(* IEC 61131-3 sources: 2026_Projet_YGO_ExcavatriceDragage/TOOLS/TEST_AUTO_CI/RESULTS/H_TREUILS_BENNE/reports (part 2) *)

(* ---- FB_BucketCloseThreshold_test.st ---- *)
(* =======================================================================
   🧪 FB_BucketCloseThreshold — seuil IHM d'ouverture benne (T262 phase B, C4)
   ───────────────────────────────────────────────────────────────────────
   Périmètre STRICT : le FB de décision en BOÎTE NOIRE. Il dérive du réglage
   IHM `ExtractionStartOpening_Pct` une DISTANCE de fermeture équivalente et
   un signal `Reached`. Il ne lit ni GVL, ni FB_Bucket, ni le cycle : aucun
   consommateur n'est testé ici (PRG_04 / FB_Bucket / FB_CycleSemiAuto
   relèvent de l'essai CODESYS et des gates mécaniques).

   ── Propriété cardinale (AC2 du contrat T262-PHASE-B) ──────────────────
   À ThresholdPct = 0, la branche est INACTIVE PAR CONSTRUCTION : `Reached`
   reste FALSE sur TOUTE la table Delta x géométrie. C'est ce qui rend la
   non-régression du comportement historique indépendante d'un MAX.

   ── Conventions ────────────────────────────────────────────────────────
   1) 1 appel `fb(...)` = 1 scan. Le FB est PUR (aucun état, aucun timer).
   2) ⚠️ Aucune assertion dans une boucle FOR/WHILE : ce build STruCpp
      SUPPRIME silencieusement les ASSERT_* du corps d'une boucle (vérifié
      dans le C++ généré). Tous les balayages sont DÉROULÉS.
   3) Tolérance 1e-6 : REAL en simple précision, littéral ST lu en double.
      Les distances attendues (p x 0,15 m) sont exactes à 1e-6 près.

   ── Géométrie de référence (valeurs persistées GVL_PERSISTENT) ─────────
   OffsetOpenM = 0,0 m · OffsetCloseM = 15,0 m · débattement = 15,0 m
   ⇒ distance équivalente = p % x 15,0 m = p x 0,15 m

   Références : DOC/WFLOW/AUDITS/DESIGN/CHALLENGE_T262_PHASE_B_SEUIL_BENNE_2026-09-21.md
                DOC/WFLOW/CONTRACTS/TASK_CONTRACT_T262_PHASE_B_BUCKET_OPENING_THRESHOLD.yaml
   ======================================================================= *)

SETUP
VAR
    FB : FB_BucketCloseThreshold;
END_VAR
END_SETUP

(* ── Groupe A · Branche INACTIVE à 0 % (AC2, AC4) ─────────────────────── *)

TEST 'TC-T262B-001 seuil 0 % : Reached FAUX sur toute la table Delta x geometrie'
    (* Balayage DEROULE. Geometrie nominale 0,0 / 15,0 m ; qualification pleine. *)
    FB.ThresholdPct := 0;
    FB.OffsetOpenM := 0.0;
    FB.OffsetCloseM := 15.0;
    FB.MeasureValid := TRUE;
    FB.IsIntermediate := TRUE;

    FB.DeltaPosition_M := 0.0;   FB();
    ASSERT_FALSE(FB.Reached, '0 % : benne ouverte (Delta = 0,0) -> Reached FAUX');
    ASSERT_FALSE(FB.Active,  '0 % : branche seuil INACTIVE');

    FB.DeltaPosition_M := 7.5;   FB();
    ASSERT_FALSE(FB.Reached, '0 % : mi-course (Delta = 7,5) -> Reached FAUX');

    FB.DeltaPosition_M := 13.0;  FB();
    ASSERT_FALSE(FB.Reached, '0 % : au seuil de la tolerance historique -> Reached FAUX');

    FB.DeltaPosition_M := 14.0;  FB();
    ASSERT_FALSE(FB.Reached, '0 % : benne fermee (Delta = 14,0) -> Reached FAUX');

    FB.DeltaPosition_M := 15.0;  FB();
    ASSERT_FALSE(FB.Reached, '0 % : sur la reference fermee -> Reached FAUX (0 % n autorise RIEN)');

    FB.DeltaPosition_M := 16.0;  FB();
    ASSERT_FALSE(FB.Reached, '0 % : sur-fermeture -> Reached FAUX');

    (* Geometrie derivee : la branche doit rester inerte quelle que soit la geometrie. *)
    FB.OffsetOpenM := -1.0;
    FB.OffsetCloseM := 20.0;
    FB.DeltaPosition_M := 19.5;  FB();
    ASSERT_FALSE(FB.Reached, '0 % : autre geometrie (debattement 21,0) -> Reached FAUX');
    ASSERT_NEAR(FB.Distance_M, 0.0, 0.000001, '0 % : distance equivalente EXACTEMENT 0,0 m');
END_TEST

TEST 'TC-T262B-002 distance equivalente : 0,15 m par pourcent (geometrie persistee)'
    (* Balayage DEROULE de p = 0 a 20 : la distance est p x 0,15 m. *)
    FB.OffsetOpenM := 0.0;
    FB.OffsetCloseM := 15.0;
    FB.MeasureValid := TRUE;
    FB.IsIntermediate := TRUE;
    FB.DeltaPosition_M := 0.0;

    FB.ThresholdPct := 0;  FB();  ASSERT_NEAR(FB.Distance_M, 0.0,  0.000001, 'p=0  -> 0,00 m');
    FB.ThresholdPct := 1;  FB();  ASSERT_NEAR(FB.Distance_M, 0.15, 0.000001, 'p=1  -> 0,15 m');
    FB.ThresholdPct := 2;  FB();  ASSERT_NEAR(FB.Distance_M, 0.30, 0.000001, 'p=2  -> 0,30 m');
    FB.ThresholdPct := 3;  FB();  ASSERT_NEAR(FB.Distance_M, 0.45, 0.000001, 'p=3  -> 0,45 m');
    FB.ThresholdPct := 4;  FB();  ASSERT_NEAR(FB.Distance_M, 0.60, 0.000001, 'p=4  -> 0,60 m');
    FB.ThresholdPct := 5;  FB();  ASSERT_NEAR(FB.Distance_M, 0.75, 0.000001, 'p=5  -> 0,75 m');
    FB.ThresholdPct := 6;  FB();  ASSERT_NEAR(FB.Distance_M, 0.90, 0.000001, 'p=6  -> 0,90 m');
    FB.ThresholdPct := 7;  FB();  ASSERT_NEAR(FB.Distance_M, 1.05, 0.000001, 'p=7  -> 1,05 m');
    FB.ThresholdPct := 8;  FB();  ASSERT_NEAR(FB.Distance_M, 1.20, 0.000001, 'p=8  -> 1,20 m (= plancher historique)');
    FB.ThresholdPct := 9;  FB();  ASSERT_NEAR(FB.Distance_M, 1.35, 0.000001, 'p=9  -> 1,35 m');
    FB.ThresholdPct := 10; FB();  ASSERT_NEAR(FB.Distance_M, 1.50, 0.000001, 'p=10 -> 1,50 m');
    FB.ThresholdPct := 13; FB();  ASSERT_NEAR(FB.Distance_M, 1.95, 0.000001, 'p=13 -> 1,95 m');
    FB.ThresholdPct := 14; FB();  ASSERT_NEAR(FB.Distance_M, 2.10, 0.000001, 'p=14 -> 2,10 m (au-dela de la tolerance 2,0)');
    FB.ThresholdPct := 19; FB();  ASSERT_NEAR(FB.Distance_M, 2.85, 0.000001, 'p=19 -> 2,85 m');
    FB.ThresholdPct := 20; FB();  ASSERT_NEAR(FB.Distance_M, 3.00, 0.000001, 'p=20 -> 3,00 m (borne haute)');
END_TEST

(* ── Groupe B · Saturation de la borne 0..20 (AC1) ────────────────────── *)

TEST 'TC-T262B-003 borne basse : seuil negatif ramene a 0 (branche INACTIVE)'
    FB.ThresholdPct := -1;
    FB.OffsetOpenM := 0.0;
    FB.OffsetCloseM := 15.0;
    FB.MeasureValid := TRUE;
    FB.IsIntermediate := TRUE;
    FB.DeltaPosition_M := 14.9;
    FB();
    ASSERT_FALSE(FB.Active, 'Seuil -1 % : branche INACTIVE');
    ASSERT_FALSE(FB.Reached, 'Seuil -1 % : Reached FAUX (aucune autorisation sur saisie hors plage)');
    ASSERT_NEAR(FB.Distance_M, 0.0, 0.000001, 'Seuil -1 % : distance ramenee a 0,0 m');
END_TEST

TEST 'TC-T262B-004 borne haute : seuil 21 ramene a 20 (jamais au-dela)'
    FB.ThresholdPct := 21;
    FB.OffsetOpenM := 0.0;
    FB.OffsetCloseM := 15.0;
    FB.MeasureValid := TRUE;
    FB.IsIntermediate := TRUE;
    FB.DeltaPosition_M := 11.5;   (* ouverture 23,3 % : hors de la plage autorisee *)
    FB();
    ASSERT_NEAR(FB.Distance_M, 3.00, 0.000001, 'Seuil 21 % : distance CLAMPEE a 3,00 m (borne 20 %)');
    ASSERT_FALSE(FB.Reached, 'Seuil 21 % : Reached FAUX a 11,5 m (la borne 20 % est respectee)');
END_TEST

TEST 'TC-T262B-005 seuil 50 (ancienne borne du contrat parent) : ramene a 20'
    FB.ThresholdPct := 50;
    FB.OffsetOpenM := 0.0;
    FB.OffsetCloseM := 15.0;
    FB.MeasureValid := TRUE;
    FB.IsIntermediate := TRUE;
    FB.DeltaPosition_M := 11.5;   (* ouverture 23,3 % : autorisee par 50 %, INTERDITE par la borne 20 % *)
    FB();
    ASSERT_NEAR(FB.Distance_M, 3.00, 0.000001, 'Seuil 50 % : distance CLAMPEE a 3,00 m (regression de borne refusee)');
    ASSERT_FALSE(FB.Reached, 'Seuil 50 % : Reached FAUX a 11,5 m -> la borne 20 % ne peut pas etre contournee');
END_TEST

(* ── Groupe C · Point de bascule au seuil (AC3) ───────────────────────── *)

TEST 'TC-T262B-006 p=10 : bascule exactement a Delta = 13,50 m (faux / vrai / vrai)'
    FB.ThresholdPct := 10;
    FB.OffsetOpenM := 0.0;
    FB.OffsetCloseM := 15.0;
    FB.MeasureValid := TRUE;
    FB.IsIntermediate := TRUE;

    FB.DeltaPosition_M := 13.49;  FB();
    ASSERT_FALSE(FB.Reached, 'p=10 : Delta = 13,49 m (ouverture 10,07 %) -> Reached FAUX');

    FB.DeltaPosition_M := 13.50;  FB();
    ASSERT_TRUE(FB.Reached, 'p=10 : Delta = 13,50 m (ouverture 10,00 %) -> Reached VRAI, egalite INCLUSE');

    FB.DeltaPosition_M := 13.51;  FB();
    ASSERT_TRUE(FB.Reached, 'p=10 : Delta = 13,51 m (ouverture 9,93 %) -> Reached VRAI');
END_TEST

TEST 'TC-T262B-007 p=19 : bascule exactement a Delta = 12,15 m'
    FB.ThresholdPct := 19;
    FB.OffsetOpenM := 0.0;
    FB.OffsetCloseM := 15.0;
    FB.MeasureValid := TRUE;
    FB.IsIntermediate := TRUE;

    FB.DeltaPosition_M := 12.14;  FB();
    ASSERT_FALSE(FB.Reached, 'p=19 : Delta = 12,14 m -> Reached FAUX');

    FB.DeltaPosition_M := 12.15;  FB();
    ASSERT_TRUE(FB.Reached, 'p=19 : Delta = 12,15 m -> Reached VRAI (egalite incluse)');

    FB.DeltaPosition_M := 12.16;  FB();
    ASSERT_TRUE(FB.Reached, 'p=19 : Delta = 12,16 m -> Reached VRAI');
END_TEST

TEST 'TC-T262B-008 p=20 (borne) : bascule exactement a Delta = 12,00 m'
    FB.ThresholdPct := 20;
    FB.OffsetOpenM := 0.0;
    FB.OffsetCloseM := 15.0;
    FB.MeasureValid := TRUE;
    FB.IsIntermediate := TRUE;

    FB.DeltaPosition_M := 11.99;  FB();
    ASSERT_FALSE(FB.Reached, 'p=20 : Delta = 11,99 m (ouverture 20,07 %) -> Reached FAUX');

    FB.DeltaPosition_M := 12.00;  FB();
    ASSERT_TRUE(FB.Reached, 'p=20 : Delta = 12,00 m (ouverture 20,00 %) -> Reached VRAI');

    FB.DeltaPosition_M := 12.01;  FB();
    ASSERT_TRUE(FB.Reached, 'p=20 : Delta = 12,01 m -> Reached VRAI');
END_TEST

(* ── Groupe D · Qualification de la mesure (AC5) ──────────────────────── *)

TEST 'TC-T262B-009 geometrie INVALIDE (OffsetOpenM >= OffsetCloseM) : jamais d autorisation'
    FB.ThresholdPct := 20;
    FB.OffsetOpenM := 15.0;      (* inversee *)
    FB.OffsetCloseM := 15.0;
    FB.MeasureValid := TRUE;
    FB.IsIntermediate := TRUE;
    FB.DeltaPosition_M := 14.9;  (* tres proche de la reference, mais geometrie inexploitable *)
    FB();
    ASSERT_FALSE(FB.Active, 'Geometrie invalide : branche seuil INACTIVE');
    ASSERT_FALSE(FB.Reached, 'Geometrie invalide : Reached FAUX (le faux 0 % ne vaut JAMAIS preuve de fermeture)');
    ASSERT_NEAR(FB.Distance_M, 0.0, 0.000001, 'Geometrie invalide : distance neutralisee a 0,0 m');
END_TEST

TEST 'TC-T262B-010 geometrie INVALIDE (OffsetOpenM > OffsetCloseM) : jamais d autorisation'
    FB.ThresholdPct := 20;
    FB.OffsetOpenM := 16.0;
    FB.OffsetCloseM := 15.0;
    FB.MeasureValid := TRUE;
    FB.IsIntermediate := TRUE;
    FB.DeltaPosition_M := 14.9;
    FB();
    ASSERT_FALSE(FB.Active, 'Geometrie inversee : branche seuil INACTIVE');
    ASSERT_FALSE(FB.Reached, 'Geometrie inversee : Reached FAUX');
    ASSERT_NEAR(FB.Distance_M, 0.0, 0.000001, 'Geometrie inversee : distance neutralisee');
END_TEST

TEST 'TC-T262B-011 MeasureValid FAUX (ActiveOffsetValid) : jamais d autorisation'
    FB.ThresholdPct := 20;
    FB.OffsetOpenM := 0.0;
    FB.OffsetCloseM := 15.0;
    FB.MeasureValid := FALSE;    (* references non fiables / defaut / puissance absente *)
    FB.IsIntermediate := TRUE;
    FB.DeltaPosition_M := 14.9;
    FB();
    ASSERT_FALSE(FB.Active, 'MeasureValid FAUX : branche seuil INACTIVE');
    ASSERT_FALSE(FB.Reached, 'MeasureValid FAUX : Reached FAUX');
END_TEST

TEST 'TC-T262B-012 IsIntermediate FAUX (mesure hors bande plausible) : jamais d autorisation'
    FB.ThresholdPct := 20;
    FB.OffsetOpenM := 0.0;
    FB.OffsetCloseM := 15.0;
    FB.MeasureValid := TRUE;
    FB.IsIntermediate := FALSE;  (* sur-fermeture / sur-ouverture : mesure non plausible *)
    FB.DeltaPosition_M := 14.9;
    FB();
    ASSERT_FALSE(FB.Active, 'IsIntermediate FAUX : branche seuil INACTIVE');
    ASSERT_FALSE(FB.Reached, 'IsIntermediate FAUX : Reached FAUX');
END_TEST

(* ── Groupe E · Pas de front : la branche reste vraie (AC9, anti-deadlock AX10) ── *)

TEST 'TC-T262B-013 p=20 : Reached reste VRAI sur 3 scans consecutifs a Delta constant'
    (* Preuve anti-deadlock : la porte AX10 ne doit pas dependre d un front present au
       scan exact d arrivee. Sans cette propriete, un geste absent au bon scan figerait
       la sortie AX10 (defaut constate et corrige par la tolerance historique). *)
    FB.ThresholdPct := 20;
    FB.OffsetOpenM := 0.0;
    FB.OffsetCloseM := 15.0;
    FB.MeasureValid := TRUE;
    FB.IsIntermediate := TRUE;
    FB.DeltaPosition_M := 12.00;

    FB();  ASSERT_TRUE(FB.Reached, 'Scan 1 : Reached VRAI');
    FB();  ASSERT_TRUE(FB.Reached, 'Scan 2 : Reached TOUJOURS VRAI (aucun front requis)');
    FB();  ASSERT_TRUE(FB.Reached, 'Scan 3 : Reached TOUJOURS VRAI');
END_TEST

TEST 'TC-T262B-014 p=20 : sortie puis retour dans la zone -> Reached de nouveau VRAI'
    FB.ThresholdPct := 20;
    FB.OffsetOpenM := 0.0;
    FB.OffsetCloseM := 15.0;
    FB.MeasureValid := TRUE;
    FB.IsIntermediate := TRUE;

    FB.DeltaPosition_M := 12.00;  FB();
    ASSERT_TRUE(FB.Reached, 'Entree dans la zone : Reached VRAI');

    FB.DeltaPosition_M := 10.00;  FB();   (* ouverture 33,3 % : hors zone *)
    ASSERT_FALSE(FB.Reached, 'Sortie de la zone : Reached FAUX');

    FB.DeltaPosition_M := 12.50;  FB();   (* geste repris, la benne se referme *)
    ASSERT_TRUE(FB.Reached, 'Retour dans la zone : Reached VRAI sans etat memorise');
END_TEST

(* ── Groupe F · Monotonie : un reglage plus grand ne resserre JAMAIS (AC4) ── *)

TEST 'TC-T262B-015 monotonie : Delta fixe, Reached VRAI pour p = seuil .. 20'
    (* Le point probatoire de la conception : augmenter le reglage ne peut JAMAIS
       rendre le critere plus strict. On se place a l ouverture 15 % (Delta = 12,75 m). *)
    FB.OffsetOpenM := 0.0;
    FB.OffsetCloseM := 15.0;
    FB.MeasureValid := TRUE;
    FB.IsIntermediate := TRUE;
    FB.DeltaPosition_M := 12.75;          (* ouverture exactement 15,00 % *)

    FB.ThresholdPct := 0;   FB();  ASSERT_FALSE(FB.Reached, 'p=0  : inerte (historique seul)');
    FB.ThresholdPct := 10;  FB();  ASSERT_FALSE(FB.Reached, 'p=10 : inerte, seuil non atteint a 15 % d ouverture');
    FB.ThresholdPct := 14;  FB();  ASSERT_FALSE(FB.Reached, 'p=14 : inerte (distance 2,10 m < 2,25 m restants)');
    FB.ThresholdPct := 15;  FB();  ASSERT_TRUE(FB.Reached,  'p=15 : BASCULE (egalite incluse)');
    FB.ThresholdPct := 16;  FB();  ASSERT_TRUE(FB.Reached,  'p=16 : VRAI (un reglage plus grand ne resserre pas)');
    FB.ThresholdPct := 20;  FB();  ASSERT_TRUE(FB.Reached,  'p=20 : VRAI (monotonie tenue jusqu a la borne)');
END_TEST

TEST 'TC-T262B-016 monotonie : Reached VRAI a p est encore VRAI a p+1 pour un Delta donne'
    (* Balayage DEROULE : Delta = 12,30 m (ouverture 18,00 %). *)
    FB.OffsetOpenM := 0.0;
    FB.OffsetCloseM := 15.0;
    FB.MeasureValid := TRUE;
    FB.IsIntermediate := TRUE;
    FB.DeltaPosition_M := 12.30;

    FB.ThresholdPct := 17;  FB();  ASSERT_FALSE(FB.Reached, 'p=17 : FAUX (distance 2,55 m > 2,70 m restants)');
    FB.ThresholdPct := 18;  FB();  ASSERT_TRUE(FB.Reached,  'p=18 : VRAI (egalite incluse)');
    FB.ThresholdPct := 19;  FB();  ASSERT_TRUE(FB.Reached,  'p=19 : VRAI');
    FB.ThresholdPct := 20;  FB();  ASSERT_TRUE(FB.Reached,  'p=20 : VRAI');
END_TEST

(* ---- FB_DriftGuard_test.st ---- *)
(* =======================================================================
   test_fb_driftguard.st — T181-18 D11 : macro TC FB_DriftGuard
   ======================================================================= *)

SETUP
VAR
    fb : FB_DriftGuard;
END_VAR
END_SETUP

TEST 'TC-P10-T181-18a Armement capture la position de reference'
    fb(Arm := FALSE, PositionM := 10.0, ToleranceM := 1.0);
    fb(Arm := TRUE, PositionM := 10.0, ToleranceM := 1.0);
    ASSERT_EQ(fb.RefPosM, 10.0, 'Reference capturee');
    ASSERT_EQ(fb.DriftM, 0.0, 'Derive nulle a la capture');
    ASSERT_FALSE(fb.Violation, 'Pas de violation');
END_TEST

TEST 'TC-P10-T181-18b Derive sous tolerance : pas de violation'
    fb(Arm := FALSE, PositionM := 10.0, ToleranceM := 1.0);
    fb(Arm := TRUE, PositionM := 10.0, ToleranceM := 1.0);
    fb(Arm := TRUE, PositionM := 10.5, ToleranceM := 1.0);
    ASSERT_EQ(fb.DriftM, 0.5, 'Derive = 0.5 m');
    ASSERT_FALSE(fb.Violation, 'Sous tolerance');
END_TEST

TEST 'TC-P10-T181-18c Derive au-dela de la tolerance : violation'
    fb(Arm := FALSE, PositionM := 10.0, ToleranceM := 1.0);
    fb(Arm := TRUE, PositionM := 10.0, ToleranceM := 1.0);
    fb(Arm := TRUE, PositionM := 11.2, ToleranceM := 1.0);
    ASSERT_TRUE(fb.Violation, 'Violation detectee au-dela de 1.0 m');
END_TEST

TEST 'TC-P10-T181-18d Desarmement puis rearmement : nouvelle reference'
    fb(Arm := FALSE, PositionM := 10.0, ToleranceM := 1.0);
    fb(Arm := TRUE, PositionM := 10.0, ToleranceM := 1.0);
    fb(Arm := FALSE, PositionM := 20.0, ToleranceM := 1.0);
    ASSERT_EQ(fb.DriftM, 0.0, 'Desarme : derive remise a zero');
    ASSERT_FALSE(fb.Violation, 'Desarme : pas de violation');
    fb(Arm := TRUE, PositionM := 20.0, ToleranceM := 1.0);
    ASSERT_EQ(fb.RefPosM, 20.0, 'Nouvelle reference a 20.0 m');
END_TEST

(* ---- FB_Safety_Winch_test.st ---- *)
(* =======================================================================
   🧪 test_fb_safety_winch.st — FB_Safety_Winch (TC-P10-001..010, 018, 036.1, 037.1, 044.1, 051.1)
   ───────────────────────────────────────────────────────────────
   Fiche : DOC/AF/AF_Partie-10_Fonction_Winch/FB_Safety_Winch_v1.0.md
   Conventions : 1 appel fb() = 1 scan ; ADVANCE_TIME(10000000) entre les
   scans pour les fronts R_TRIG ; hex décrit en décimal (bit 0 = 1, bit 15 = 32768).
   Masque PowerCutOff = 16#2F84 = bits 2,7,8,9,10,11,13 (décimal 12164).
   Masque SafeStop SyncEnable=TRUE  = 16#FF9F ; SyncEnable=FALSE = 16#FF97 (exclut bit3).
   ======================================================================= *)

SETUP
VAR
    fb : FB_Safety_Winch;
END_VAR
END_SETUP

(* ── Remise à zéro commune : pulse Enable+Reset, puis Reset retombé ── *)

TEST 'TC-P10-001 Meca A : derive >5.0m a l arret (joystick neutre) -> SafeStop + PowerCutOff'
    (* Scan 1 : Enable=TRUE, regime nominal, joystick neutre, contacteurs+frein confirmes coupes *)
    fb(Enable := TRUE, Reset := FALSE, SyncEnable := FALSE,
       PowerContactorEngaged := TRUE, JoystickOnline := TRUE, JoystickOperational := TRUE,
       HeartbeatIhmOk := TRUE, EncoderAvailable := TRUE, PhaseRotationOk := TRUE,
       TopPositionSensor := TRUE, FwdRevSpeedFeedbackOff := TRUE, BrakeFeedback := FALSE,
       JoystickYNeutral := TRUE, BenneHoldStillActive := FALSE, InReferencingMode := FALSE,
       CablePosM := 0.0, CfgCableLimitDescentM := -20.0, Homed := TRUE, TopLimitM := 8.5);
    ADVANCE_TIME(10000000);
    (* Scan 2 : regime etabli, Meca A arme (RefPosM capture a 0.0) *)
    fb(Enable := TRUE, Reset := FALSE, SyncEnable := FALSE,
       PowerContactorEngaged := TRUE, JoystickOnline := TRUE, JoystickOperational := TRUE,
       HeartbeatIhmOk := TRUE, EncoderAvailable := TRUE, PhaseRotationOk := TRUE,
       TopPositionSensor := TRUE, FwdRevSpeedFeedbackOff := TRUE, BrakeFeedback := FALSE,
       JoystickYNeutral := TRUE, BenneHoldStillActive := FALSE, InReferencingMode := FALSE,
       CablePosM := 0.0, CfgCableLimitDescentM := -20.0, Homed := TRUE, TopLimitM := 8.5);
    ASSERT_FALSE(fb.SafeStop, 'Nominal : pas de SafeStop');
    ASSERT_FALSE(fb.PowerCutOff, 'Nominal : pas de PowerCutOff');
    ASSERT_FALSE(fb.Fault.Error, 'Nominal : pas d erreur');
    (* Scan 3 : derive injectee > 5.0m (mono-canal position) - MES 2026-09-04 : seuil 2.0->5.0m *)
    ADVANCE_TIME(10000000);
    fb(Enable := TRUE, Reset := FALSE, SyncEnable := FALSE,
       PowerContactorEngaged := TRUE, JoystickOnline := TRUE, JoystickOperational := TRUE,
       HeartbeatIhmOk := TRUE, EncoderAvailable := TRUE, PhaseRotationOk := TRUE,
       TopPositionSensor := TRUE, FwdRevSpeedFeedbackOff := TRUE, BrakeFeedback := FALSE,
       JoystickYNeutral := TRUE, BenneHoldStillActive := FALSE, InReferencingMode := FALSE,
       CablePosM := 6.0, CfgCableLimitDescentM := -20.0, Homed := TRUE, TopLimitM := 8.5);
    ASSERT_TRUE(fb.SafeStop, 'Derive >5.0m -> SafeStop');
    ASSERT_TRUE(fb.PowerCutOff, 'Derive >5.0m -> PowerCutOff (bit7 dans masque 16#2F84)');
    ASSERT_TRUE(fb.Fault.Error, 'Derive >5.0m -> Error');
    ASSERT_TRUE(fb.Fault.Latched, 'Meca A latchee (defaut a acquitter)');
END_TEST

TEST 'TC-P10-054 T288 : retour collectif au repos sous commande 3s -> SafeStop seul'
    (* Cas terrain 14/09 : commande active, frein ouvert, retour collectif
       tous contacteurs retombes et codeur immobile. *)
    fb(Enable := TRUE, Reset := FALSE, SyncEnable := FALSE,
       PowerContactorEngaged := TRUE, JoystickOnline := TRUE, JoystickOperational := TRUE,
       HeartbeatIhmOk := TRUE, EncoderAvailable := TRUE, PhaseRotationOk := TRUE,
       TopPositionSensor := TRUE, FwdRevSpeedFeedbackOff := TRUE, BrakeFeedback := FALSE,
       JoystickYNeutral := TRUE, BenneHoldStillActive := FALSE, InReferencingMode := FALSE,
       CablePosM := 0.0, CfgCableLimitDescentM := -20.0, Homed := TRUE, TopLimitM := 8.5);
    (* Attendre la fenetre de reference existante avant d armer la surveillance. *)
    ADVANCE_TIME(3000000000);
    fb(Enable := TRUE, Reset := FALSE, SyncEnable := FALSE,
       PowerContactorEngaged := TRUE, JoystickOnline := TRUE, JoystickOperational := TRUE,
       HeartbeatIhmOk := TRUE, EncoderAvailable := TRUE, PhaseRotationOk := TRUE,
       TopPositionSensor := TRUE, FwdRevSpeedFeedbackOff := TRUE, BrakeFeedback := FALSE,
       JoystickYNeutral := TRUE, BenneHoldStillActive := FALSE, InReferencingMode := FALSE,
       CablePosM := 0.0, CfgCableLimitDescentM := -20.0, Homed := TRUE, TopLimitM := 8.5);
    ADVANCE_TIME(10000000);
    fb(Enable := TRUE, Reset := FALSE, SyncEnable := FALSE,
       PowerContactorEngaged := TRUE, JoystickOnline := TRUE, JoystickOperational := TRUE,
       HeartbeatIhmOk := TRUE, EncoderAvailable := TRUE, PhaseRotationOk := TRUE,
       TopPositionSensor := TRUE, FwdRevSpeedFeedbackOff := TRUE, BrakeFeedback := TRUE,
       JoystickYNeutral := FALSE, BenneHoldStillActive := FALSE, InReferencingMode := FALSE,
       CablePosM := 0.0, CfgCableLimitDescentM := -20.0, Homed := TRUE, TopLimitM := 8.5,
       ReqAscent := TRUE, ReqDescend := FALSE, MovementCommanded := TRUE);
    ASSERT_FALSE(fb.SafeStop, 'Avant 3s : pas de SafeStop');
    ADVANCE_TIME(3000000000);
    fb(Enable := TRUE, Reset := FALSE, SyncEnable := FALSE,
       PowerContactorEngaged := TRUE, JoystickOnline := TRUE, JoystickOperational := TRUE,
       HeartbeatIhmOk := TRUE, EncoderAvailable := TRUE, PhaseRotationOk := TRUE,
       TopPositionSensor := TRUE, FwdRevSpeedFeedbackOff := TRUE, BrakeFeedback := TRUE,
       JoystickYNeutral := FALSE, BenneHoldStillActive := FALSE, InReferencingMode := FALSE,
       CablePosM := 0.0, CfgCableLimitDescentM := -20.0, Homed := TRUE, TopLimitM := 8.5,
       ReqAscent := TRUE, ReqDescend := FALSE, MovementCommanded := TRUE);
    ASSERT_TRUE(fb.SafeStop, 'Retour collectif au repos + aucun mouvement 3s -> SafeStop');
    ASSERT_FALSE(fb.PowerCutOff, 'T288 -> SafeStop seul, sans PowerCutOff');
    ASSERT_TRUE(fb.Fault.Error, 'T288 -> ErrorID 16 actif');
END_TEST

TEST 'TC-P10-055 T288 : retour collectif engage sous commande 3s -> SafeStop seul'
    (* Variante historique : au moins un contacteur confirme mais le codeur reste immobile. *)
    fb(Enable := TRUE, Reset := FALSE, SyncEnable := FALSE,
       PowerContactorEngaged := TRUE, JoystickOnline := TRUE, JoystickOperational := TRUE,
       HeartbeatIhmOk := TRUE, EncoderAvailable := TRUE, PhaseRotationOk := TRUE,
       TopPositionSensor := TRUE, FwdRevSpeedFeedbackOff := TRUE, BrakeFeedback := FALSE,
       JoystickYNeutral := TRUE, BenneHoldStillActive := FALSE, InReferencingMode := FALSE,
       CablePosM := 0.0, CfgCableLimitDescentM := -20.0, Homed := TRUE, TopLimitM := 8.5);
    ADVANCE_TIME(3000000000);
    fb(Enable := TRUE, Reset := FALSE, SyncEnable := FALSE,
       PowerContactorEngaged := TRUE, JoystickOnline := TRUE, JoystickOperational := TRUE,
       HeartbeatIhmOk := TRUE, EncoderAvailable := TRUE, PhaseRotationOk := TRUE,
       TopPositionSensor := TRUE, FwdRevSpeedFeedbackOff := TRUE, BrakeFeedback := FALSE,
       JoystickYNeutral := TRUE, BenneHoldStillActive := FALSE, InReferencingMode := FALSE,
       CablePosM := 0.0, CfgCableLimitDescentM := -20.0, Homed := TRUE, TopLimitM := 8.5);
    ADVANCE_TIME(10000000);
    fb(Enable := TRUE, Reset := FALSE, SyncEnable := FALSE,
       PowerContactorEngaged := TRUE, JoystickOnline := TRUE, JoystickOperational := TRUE,
       HeartbeatIhmOk := TRUE, EncoderAvailable := TRUE, PhaseRotationOk := TRUE,
       TopPositionSensor := TRUE, FwdRevSpeedFeedbackOff := FALSE, BrakeFeedback := TRUE,
       JoystickYNeutral := FALSE, BenneHoldStillActive := FALSE, InReferencingMode := FALSE,
       CablePosM := 0.0, CfgCableLimitDescentM := -20.0, Homed := TRUE, TopLimitM := 8.5,
       ReqAscent := TRUE, ReqDescend := FALSE, MovementCommanded := TRUE);
    ASSERT_FALSE(fb.SafeStop, 'Avant 3s : pas de SafeStop');
    ADVANCE_TIME(3000000000);
    fb(Enable := TRUE, Reset := FALSE, SyncEnable := FALSE,
       PowerContactorEngaged := TRUE, JoystickOnline := TRUE, JoystickOperational := TRUE,
       HeartbeatIhmOk := TRUE, EncoderAvailable := TRUE, PhaseRotationOk := TRUE,
       TopPositionSensor := TRUE, FwdRevSpeedFeedbackOff := FALSE, BrakeFeedback := TRUE,
       JoystickYNeutral := FALSE, BenneHoldStillActive := FALSE, InReferencingMode := FALSE,
       CablePosM := 0.0, CfgCableLimitDescentM := -20.0, Homed := TRUE, TopLimitM := 8.5,
       ReqAscent := TRUE, ReqDescend := FALSE, MovementCommanded := TRUE);
    ASSERT_TRUE(fb.SafeStop, 'Retour collectif engage + aucun mouvement 3s -> SafeStop');
    ASSERT_FALSE(fb.PowerCutOff, 'T288 historique -> SafeStop seul, sans PowerCutOff');
END_TEST

TEST 'TC-P10-002 Meca B : non confirmation arret 3s -> SafeStop + PowerCutOff'
    (* Scan 1 : regime nominal *)
    fb(Enable := TRUE, Reset := FALSE, SyncEnable := FALSE,
       PowerContactorEngaged := TRUE, JoystickOnline := TRUE, JoystickOperational := TRUE,
       HeartbeatIhmOk := TRUE, EncoderAvailable := TRUE, PhaseRotationOk := TRUE,
       TopPositionSensor := TRUE, FwdRevSpeedFeedbackOff := TRUE, BrakeFeedback := FALSE,
       JoystickYNeutral := TRUE, BenneHoldStillActive := FALSE, InReferencingMode := FALSE,
       CablePosM := 0.0, CfgCableLimitDescentM := -20.0, Homed := TRUE, TopLimitM := 8.5);
    ADVANCE_TIME(10000000);
    (* Scan 2 : joystick neutre mais contacteurs NON confirmes retombes (FwdRevSpeedFeedbackOff=FALSE) *)
    fb(Enable := TRUE, Reset := FALSE, SyncEnable := FALSE,
       PowerContactorEngaged := TRUE, JoystickOnline := TRUE, JoystickOperational := TRUE,
       HeartbeatIhmOk := TRUE, EncoderAvailable := TRUE, PhaseRotationOk := TRUE,
       TopPositionSensor := TRUE, FwdRevSpeedFeedbackOff := FALSE, BrakeFeedback := FALSE,
       JoystickYNeutral := TRUE, BenneHoldStillActive := FALSE, InReferencingMode := FALSE,
       CablePosM := 0.0, CfgCableLimitDescentM := -20.0, Homed := TRUE, TopLimitM := 8.5);
    ASSERT_FALSE(fb.PowerCutOff, 'Avant 3s : pas encore de PowerCutOff');
    (* Scan 3 : apres PostRampTimeout=3s -> Meca B latchee *)
    ADVANCE_TIME(3000000000);
    fb(Enable := TRUE, Reset := FALSE, SyncEnable := FALSE,
       PowerContactorEngaged := TRUE, JoystickOnline := TRUE, JoystickOperational := TRUE,
       HeartbeatIhmOk := TRUE, EncoderAvailable := TRUE, PhaseRotationOk := TRUE,
       TopPositionSensor := TRUE, FwdRevSpeedFeedbackOff := FALSE, BrakeFeedback := FALSE,
       JoystickYNeutral := TRUE, BenneHoldStillActive := FALSE, InReferencingMode := FALSE,
       CablePosM := 0.0, CfgCableLimitDescentM := -20.0, Homed := TRUE, TopLimitM := 8.5);
    ASSERT_TRUE(fb.SafeStop, 'Non confirmation arret 3s -> SafeStop');
    ASSERT_TRUE(fb.PowerCutOff, 'Non confirmation arret 3s -> PowerCutOff (bit8 dans masque)');
    ASSERT_TRUE(fb.Fault.Error, 'Meca B -> Error');
END_TEST

TEST 'TC-P10-018 ContactorStuck : contacteur colle -> ContactorStuck + SafeStop + PowerCutOff (action, pas seulement diagnostic)'
    (* (adapte depuis TC-P10-018 FB_Winch, T181-02/03 AC5) : FB_Safety_Winch est le producteur
       UNIQUE de ContactorStuck. Le TC prouve l'ACTION de securite (SafeStop + PowerCutOff),
       pas seulement l'etat diagnostic. *)
    (* Scan 1 : regime nominal *)
    fb(Enable := TRUE, Reset := FALSE, SyncEnable := FALSE,
       PowerContactorEngaged := TRUE, JoystickOnline := TRUE, JoystickOperational := TRUE,
       HeartbeatIhmOk := TRUE, EncoderAvailable := TRUE, PhaseRotationOk := TRUE,
       TopPositionSensor := TRUE, FwdRevSpeedFeedbackOff := TRUE, BrakeFeedback := FALSE,
       JoystickYNeutral := TRUE, BenneHoldStillActive := FALSE, InReferencingMode := FALSE,
       CablePosM := 0.0, CfgCableLimitDescentM := -20.0, Homed := TRUE, TopLimitM := 8.5);
    ADVANCE_TIME(10000000);
    (* Scan 2 : joystick neutre mais contacteurs NON retombes (FwdRevSpeedFeedbackOff=FALSE) *)
    fb(Enable := TRUE, Reset := FALSE, SyncEnable := FALSE,
       PowerContactorEngaged := TRUE, JoystickOnline := TRUE, JoystickOperational := TRUE,
       HeartbeatIhmOk := TRUE, EncoderAvailable := TRUE, PhaseRotationOk := TRUE,
       TopPositionSensor := TRUE, FwdRevSpeedFeedbackOff := FALSE, BrakeFeedback := FALSE,
       JoystickYNeutral := TRUE, BenneHoldStillActive := FALSE, InReferencingMode := FALSE,
       CablePosM := 0.0, CfgCableLimitDescentM := -20.0, Homed := TRUE, TopLimitM := 8.5);
    ASSERT_FALSE(fb.ContactorStuck, 'Avant 3s : pas encore de ContactorStuck');
    ASSERT_FALSE(fb.PowerCutOff, 'Avant 3s : pas encore de PowerCutOff');
    (* Scan 3 : apres PostRampTimeout=3s -> ContactorStuck + SafeStop + PowerCutOff *)
    ADVANCE_TIME(3000000000);
    fb(Enable := TRUE, Reset := FALSE, SyncEnable := FALSE,
       PowerContactorEngaged := TRUE, JoystickOnline := TRUE, JoystickOperational := TRUE,
       HeartbeatIhmOk := TRUE, EncoderAvailable := TRUE, PhaseRotationOk := TRUE,
       TopPositionSensor := TRUE, FwdRevSpeedFeedbackOff := FALSE, BrakeFeedback := FALSE,
       JoystickYNeutral := TRUE, BenneHoldStillActive := FALSE, InReferencingMode := FALSE,
       CablePosM := 0.0, CfgCableLimitDescentM := -20.0, Homed := TRUE, TopLimitM := 8.5);
    ASSERT_TRUE(fb.ContactorStuck, 'Contacteur colle 3s -> ContactorStuck=TRUE');
    ASSERT_TRUE(fb.SafeStop, 'Contacteur colle -> SafeStop (action)');
    ASSERT_TRUE(fb.PowerCutOff, 'Contacteur colle -> PowerCutOff (action)');
    ASSERT_TRUE(fb.Fault.Error, 'Contacteur colle -> Error');
END_TEST

TEST 'TC-P10-003 Meca C : glissement M1 >2.0m pendant maintien benne -> SafeStop + PowerCutOff'
    (* Scan 1 : regime nominal *)
    fb(Enable := TRUE, Reset := FALSE, SyncEnable := FALSE,
       PowerContactorEngaged := TRUE, JoystickOnline := TRUE, JoystickOperational := TRUE,
       HeartbeatIhmOk := TRUE, EncoderAvailable := TRUE, PhaseRotationOk := TRUE,
       TopPositionSensor := TRUE, FwdRevSpeedFeedbackOff := TRUE, BrakeFeedback := FALSE,
       JoystickYNeutral := TRUE, BenneHoldStillActive := FALSE, InReferencingMode := FALSE,
       CablePosM := 0.0, CfgCableLimitDescentM := -20.0, Homed := TRUE, TopLimitM := 8.5);
    ADVANCE_TIME(10000000);
    (* Scan 2 : BenneHoldStillActive=TRUE -> Meca C arme (RefPosM capture a 0.0) *)
    fb(Enable := TRUE, Reset := FALSE, SyncEnable := FALSE,
       PowerContactorEngaged := TRUE, JoystickOnline := TRUE, JoystickOperational := TRUE,
       HeartbeatIhmOk := TRUE, EncoderAvailable := TRUE, PhaseRotationOk := TRUE,
       TopPositionSensor := TRUE, FwdRevSpeedFeedbackOff := TRUE, BrakeFeedback := FALSE,
       JoystickYNeutral := TRUE, BenneHoldStillActive := TRUE, InReferencingMode := FALSE,
       CablePosM := 0.0, CfgCableLimitDescentM := -20.0, Homed := TRUE, TopLimitM := 8.5);
    (* Scan 3 : derive M1 > 2.0m pendant maintien *)
    ADVANCE_TIME(10000000);
    fb(Enable := TRUE, Reset := FALSE, SyncEnable := FALSE,
       PowerContactorEngaged := TRUE, JoystickOnline := TRUE, JoystickOperational := TRUE,
       HeartbeatIhmOk := TRUE, EncoderAvailable := TRUE, PhaseRotationOk := TRUE,
       TopPositionSensor := TRUE, FwdRevSpeedFeedbackOff := TRUE, BrakeFeedback := FALSE,
       JoystickYNeutral := TRUE, BenneHoldStillActive := TRUE, InReferencingMode := FALSE,
       CablePosM := 3.0, CfgCableLimitDescentM := -20.0, Homed := TRUE, TopLimitM := 8.5);
    ASSERT_TRUE(fb.SafeStop, 'Glissement M1 >2.0m -> SafeStop');
    ASSERT_TRUE(fb.PowerCutOff, 'Glissement M1 >2.0m -> PowerCutOff (bit9 dans masque)');
    ASSERT_TRUE(fb.Fault.Error, 'Meca C -> Error');
END_TEST

TEST 'TC-P10-004 Meca D : capteur haut sans arret 3s -> SafeStop (immediat) puis PowerCutOff (3s)'
    (* Scan 1 : regime nominal *)
    fb(Enable := TRUE, Reset := FALSE, SyncEnable := FALSE,
       PowerContactorEngaged := TRUE, JoystickOnline := TRUE, JoystickOperational := TRUE,
       HeartbeatIhmOk := TRUE, EncoderAvailable := TRUE, PhaseRotationOk := TRUE,
       TopPositionSensor := TRUE, FwdRevSpeedFeedbackOff := TRUE, BrakeFeedback := FALSE,
       JoystickYNeutral := TRUE, BenneHoldStillActive := FALSE, InReferencingMode := FALSE,
       CablePosM := 0.0, CfgCableLimitDescentM := -20.0, Homed := TRUE, TopLimitM := 8.5);
    ADVANCE_TIME(10000000);
    (* Scan 2 : capteur haut atteint (TopPositionSensor=FALSE) + contacteurs non retombes.
       Cause 5 (fin de course haut) -> AscentPermit=FALSE (bit5 hors masque SafeStop 16#FF97) ;
       SafeStop/PowerCutOff viennent de Meca D (bit11) apres 3s. *)
    fb(Enable := TRUE, Reset := FALSE, SyncEnable := FALSE,
       PowerContactorEngaged := TRUE, JoystickOnline := TRUE, JoystickOperational := TRUE,
       HeartbeatIhmOk := TRUE, EncoderAvailable := TRUE, PhaseRotationOk := TRUE,
       TopPositionSensor := FALSE, FwdRevSpeedFeedbackOff := FALSE, BrakeFeedback := FALSE,
       JoystickYNeutral := TRUE, BenneHoldStillActive := FALSE, InReferencingMode := FALSE,
       CablePosM := 0.0, CfgCableLimitDescentM := -20.0, Homed := TRUE, TopLimitM := 8.5);
    ASSERT_FALSE(fb.AscentPermit, 'Capteur haut atteint -> AscentPermit=FALSE (cause 5)');
    ASSERT_FALSE(fb.SafeStop, 'Avant 3s : Meca D pas encore latchee -> pas de SafeStop');
    ASSERT_FALSE(fb.PowerCutOff, 'Avant 3s : Meca D pas encore latchee -> pas de PowerCutOff');
    (* Scan 3 : apres PostRampTimeout=3s -> Meca D latchee -> SafeStop + PowerCutOff *)
    ADVANCE_TIME(3000000000);
    fb(Enable := TRUE, Reset := FALSE, SyncEnable := FALSE,
       PowerContactorEngaged := TRUE, JoystickOnline := TRUE, JoystickOperational := TRUE,
       HeartbeatIhmOk := TRUE, EncoderAvailable := TRUE, PhaseRotationOk := TRUE,
       TopPositionSensor := FALSE, FwdRevSpeedFeedbackOff := FALSE, BrakeFeedback := FALSE,
       JoystickYNeutral := TRUE, BenneHoldStillActive := FALSE, InReferencingMode := FALSE,
       CablePosM := 0.0, CfgCableLimitDescentM := -20.0, Homed := TRUE, TopLimitM := 8.5);
    ASSERT_TRUE(fb.SafeStop, 'Capteur haut sans arret 3s -> SafeStop (Meca D bit11)');
    ASSERT_TRUE(fb.PowerCutOff, 'Capteur haut sans arret 3s -> PowerCutOff (bit11 dans masque)');
    ASSERT_TRUE(fb.Fault.Error, 'Meca D -> Error');
END_TEST

TEST 'TC-P10-005 Meca E bit12 : ecart >2.5m -> SafeStop SEUL (pas PowerCutOff)'
    (* BypassMecaA=TRUE isole Meca E : l armement Meca A est desormais base sur le retour
       mecanique, pas sur JoystickYNeutral. Seul Meca E (bit12) doit se declencher. *)
    (* Scan 1 : regime nominal avec SyncEnable=TRUE *)
    fb(Enable := TRUE, Reset := FALSE, SyncEnable := TRUE,
       PowerContactorEngaged := TRUE, JoystickOnline := TRUE, JoystickOperational := TRUE,
       HeartbeatIhmOk := TRUE, EncoderAvailable := TRUE, PhaseRotationOk := TRUE,
       TopPositionSensor := TRUE, FwdRevSpeedFeedbackOff := TRUE, BrakeFeedback := FALSE,
       JoystickYNeutral := FALSE, BenneHoldStillActive := FALSE, BenneBusy := FALSE,
       OtherWinchInhibited := FALSE, InReferencingMode := FALSE, BypassMecaA := TRUE,
       CablePosM := 0.0, ExpectedOtherWinchPosM := 0.0, CfgCableLimitDescentM := -20.0,
       Homed := TRUE, TopLimitM := 8.5);
    ADVANCE_TIME(10000000);
    (* Scan 2 : ecart M1/M2 > CriticalSyncToleranceM=2.5m *)
    fb(Enable := TRUE, Reset := FALSE, SyncEnable := TRUE,
       PowerContactorEngaged := TRUE, JoystickOnline := TRUE, JoystickOperational := TRUE,
       HeartbeatIhmOk := TRUE, EncoderAvailable := TRUE, PhaseRotationOk := TRUE,
       TopPositionSensor := TRUE, FwdRevSpeedFeedbackOff := TRUE, BrakeFeedback := FALSE,
       JoystickYNeutral := FALSE, BenneHoldStillActive := FALSE, BenneBusy := FALSE,
       OtherWinchInhibited := FALSE, InReferencingMode := FALSE, BypassMecaA := TRUE,
       CablePosM := 3.0, ExpectedOtherWinchPosM := 0.0, CfgCableLimitDescentM := -20.0,
       Homed := TRUE, TopLimitM := 8.5);
    ASSERT_TRUE(fb.SafeStop, 'Ecart critique -> SafeStop (bit12 dans masque SafeStop)');
    ASSERT_FALSE(fb.PowerCutOff, 'Ecart critique bit12 -> PAS de PowerCutOff (bit12 hors masque 16#2F84)');
    ASSERT_TRUE(fb.Fault.Error, 'Meca E bit12 -> Error');
END_TEST

TEST 'TC-P10-006 Meca E bit13 : bit12 non confirme 3s -> escalade PowerCutOff'
    (* JoystickYNeutral=FALSE pour isoler Meca E (evite Meca A dans le masque PowerCutOff). *)
    (* Scan 1 : regime nominal avec SyncEnable=TRUE, ecart critique -> bit12 latche *)
    fb(Enable := TRUE, Reset := FALSE, SyncEnable := TRUE,
       PowerContactorEngaged := TRUE, JoystickOnline := TRUE, JoystickOperational := TRUE,
       HeartbeatIhmOk := TRUE, EncoderAvailable := TRUE, PhaseRotationOk := TRUE,
       TopPositionSensor := TRUE, FwdRevSpeedFeedbackOff := TRUE, BrakeFeedback := FALSE,
       JoystickYNeutral := FALSE, BenneHoldStillActive := FALSE, BenneBusy := FALSE,
       OtherWinchInhibited := FALSE, InReferencingMode := FALSE,
       CablePosM := 3.0, ExpectedOtherWinchPosM := 0.0, CfgCableLimitDescentM := -20.0,
       Homed := TRUE, TopLimitM := 8.5);
    ADVANCE_TIME(10000000);
    (* Scan 2 : bit12 latche, contacteurs non retombes -> TonMecaE arme *)
    fb(Enable := TRUE, Reset := FALSE, SyncEnable := TRUE,
       PowerContactorEngaged := TRUE, JoystickOnline := TRUE, JoystickOperational := TRUE,
       HeartbeatIhmOk := TRUE, EncoderAvailable := TRUE, PhaseRotationOk := TRUE,
       TopPositionSensor := TRUE, FwdRevSpeedFeedbackOff := FALSE, BrakeFeedback := FALSE,
       JoystickYNeutral := FALSE, BenneHoldStillActive := FALSE, BenneBusy := FALSE,
       OtherWinchInhibited := FALSE, InReferencingMode := FALSE,
       CablePosM := 3.0, ExpectedOtherWinchPosM := 0.0, CfgCableLimitDescentM := -20.0,
       Homed := TRUE, TopLimitM := 8.5);
    ASSERT_FALSE(fb.PowerCutOff, 'Avant 3s : bit12 seul -> pas de PowerCutOff');
    (* Scan 3 : apres PostRampTimeout=3s -> escalade bit13 -> PowerCutOff *)
    ADVANCE_TIME(3000000000);
    fb(Enable := TRUE, Reset := FALSE, SyncEnable := TRUE,
       PowerContactorEngaged := TRUE, JoystickOnline := TRUE, JoystickOperational := TRUE,
       HeartbeatIhmOk := TRUE, EncoderAvailable := TRUE, PhaseRotationOk := TRUE,
       TopPositionSensor := TRUE, FwdRevSpeedFeedbackOff := FALSE, BrakeFeedback := FALSE,
       JoystickYNeutral := FALSE, BenneHoldStillActive := FALSE, BenneBusy := FALSE,
       OtherWinchInhibited := FALSE, InReferencingMode := FALSE,
       CablePosM := 3.0, ExpectedOtherWinchPosM := 0.0, CfgCableLimitDescentM := -20.0,
       Homed := TRUE, TopLimitM := 8.5);
    ASSERT_TRUE(fb.PowerCutOff, 'Escalade bit13 -> PowerCutOff (bit13 dans masque 16#2F84)');
    ASSERT_TRUE(fb.Fault.Error, 'Meca E escalade -> Error');
END_TEST

TEST 'TC-P10-007 Meca F : sens mesure oppose a la commande 500ms -> SafeStop SEUL'
    (* Scan 1 : regime nominal *)
    fb(Enable := TRUE, Reset := FALSE, SyncEnable := FALSE,
       PowerContactorEngaged := TRUE, JoystickOnline := TRUE, JoystickOperational := TRUE,
       HeartbeatIhmOk := TRUE, EncoderAvailable := TRUE, PhaseRotationOk := TRUE,
       TopPositionSensor := TRUE, FwdRevSpeedFeedbackOff := TRUE, BrakeFeedback := FALSE,
       JoystickYNeutral := TRUE, BenneHoldStillActive := FALSE, InReferencingMode := FALSE,
       CablePosM := 0.0, CfgCableLimitDescentM := -20.0, Homed := TRUE, TopLimitM := 8.5);
    ADVANCE_TIME(10000000);
    (* Scan 2 : commande montee (Direction=1) mais vitesse mesuree negative *)
    fb(Enable := TRUE, Reset := FALSE, SyncEnable := FALSE,
       PowerContactorEngaged := TRUE, JoystickOnline := TRUE, JoystickOperational := TRUE,
       HeartbeatIhmOk := TRUE, EncoderAvailable := TRUE, PhaseRotationOk := TRUE,
       TopPositionSensor := TRUE, FwdRevSpeedFeedbackOff := TRUE, BrakeFeedback := FALSE,
       JoystickYNeutral := TRUE, BenneHoldStillActive := FALSE, InReferencingMode := FALSE,
       CablePosM := 0.0, CfgCableLimitDescentM := -20.0, Homed := TRUE, TopLimitM := 8.5,
       ReqAscent := TRUE, ReqDescend := FALSE, MovementCommanded := TRUE, MeasuredSpeedValid := TRUE,
       MeasuredSpeedSignedMps := -0.1);
    ASSERT_FALSE(fb.PowerCutOff, 'Avant 500ms : pas de PowerCutOff');
    (* Scan 3 : apres OppositeDirectionTimeout=500ms -> Meca F latchee *)
    ADVANCE_TIME(500000000);
    fb(Enable := TRUE, Reset := FALSE, SyncEnable := FALSE,
       PowerContactorEngaged := TRUE, JoystickOnline := TRUE, JoystickOperational := TRUE,
       HeartbeatIhmOk := TRUE, EncoderAvailable := TRUE, PhaseRotationOk := TRUE,
       TopPositionSensor := TRUE, FwdRevSpeedFeedbackOff := TRUE, BrakeFeedback := FALSE,
       JoystickYNeutral := TRUE, BenneHoldStillActive := FALSE, InReferencingMode := FALSE,
       CablePosM := 0.0, CfgCableLimitDescentM := -20.0, Homed := TRUE, TopLimitM := 8.5,
       ReqAscent := TRUE, ReqDescend := FALSE, MovementCommanded := TRUE, MeasuredSpeedValid := TRUE,
       MeasuredSpeedSignedMps := -0.1);
    ASSERT_TRUE(fb.SafeStop, 'Sens oppose 500ms -> SafeStop (bit14 dans masque)');
    ASSERT_FALSE(fb.PowerCutOff, 'Sens oppose -> PAS de PowerCutOff (bit14 hors masque 16#2F84)');
    ASSERT_TRUE(fb.Fault.Error, 'Meca F -> Error');
END_TEST

TEST 'TC-P10-008 Meca G : vitesse nulle malgre commande 3s -> SafeStop SEUL'
    (* Scan 1 : regime nominal *)
    fb(Enable := TRUE, Reset := FALSE, SyncEnable := FALSE,
       PowerContactorEngaged := TRUE, JoystickOnline := TRUE, JoystickOperational := TRUE,
       HeartbeatIhmOk := TRUE, EncoderAvailable := TRUE, PhaseRotationOk := TRUE,
       TopPositionSensor := TRUE, FwdRevSpeedFeedbackOff := TRUE, BrakeFeedback := FALSE,
       JoystickYNeutral := TRUE, BenneHoldStillActive := FALSE, InReferencingMode := FALSE,
       CablePosM := 0.0, CfgCableLimitDescentM := -20.0, Homed := TRUE, TopLimitM := 8.5);
    ADVANCE_TIME(10000000);
    (* Scan 2 : commande montee mais vitesse nulle *)
    fb(Enable := TRUE, Reset := FALSE, SyncEnable := FALSE,
       PowerContactorEngaged := TRUE, JoystickOnline := TRUE, JoystickOperational := TRUE,
       HeartbeatIhmOk := TRUE, EncoderAvailable := TRUE, PhaseRotationOk := TRUE,
       TopPositionSensor := TRUE, FwdRevSpeedFeedbackOff := TRUE, BrakeFeedback := FALSE,
       JoystickYNeutral := TRUE, BenneHoldStillActive := FALSE, InReferencingMode := FALSE,
       CablePosM := 0.0, CfgCableLimitDescentM := -20.0, Homed := TRUE, TopLimitM := 8.5,
       ReqAscent := TRUE, ReqDescend := FALSE, MovementCommanded := TRUE, MeasuredSpeedValid := TRUE,
       MeasuredSpeedSignedMps := 0.0);
    ASSERT_FALSE(fb.PowerCutOff, 'Avant 3s : pas de PowerCutOff');
    (* Scan 3 : apres NoMovementTimeout=3s -> Meca G latchee *)
    ADVANCE_TIME(3000000000);
    fb(Enable := TRUE, Reset := FALSE, SyncEnable := FALSE,
       PowerContactorEngaged := TRUE, JoystickOnline := TRUE, JoystickOperational := TRUE,
       HeartbeatIhmOk := TRUE, EncoderAvailable := TRUE, PhaseRotationOk := TRUE,
       TopPositionSensor := TRUE, FwdRevSpeedFeedbackOff := TRUE, BrakeFeedback := FALSE,
       JoystickYNeutral := TRUE, BenneHoldStillActive := FALSE, InReferencingMode := FALSE,
       CablePosM := 0.0, CfgCableLimitDescentM := -20.0, Homed := TRUE, TopLimitM := 8.5,
       ReqAscent := TRUE, ReqDescend := FALSE, MovementCommanded := TRUE, MeasuredSpeedValid := TRUE,
       MeasuredSpeedSignedMps := 0.0);
    ASSERT_TRUE(fb.SafeStop, 'Absence mouvement 3s -> SafeStop (bit15 dans masque)');
    ASSERT_FALSE(fb.PowerCutOff, 'Absence mouvement -> PAS de PowerCutOff (bit15 hors masque 16#2F84)');
    ASSERT_TRUE(fb.Fault.Error, 'Meca G -> Error');
END_TEST

TEST 'TC-P10-009 Masque PowerCutOff : bit2 (surchauffe moteur) coupe, bit14 (sens oppose) ne coupe pas'
    (* Scan 1 : regime nominal *)
    fb(Enable := TRUE, Reset := FALSE, SyncEnable := FALSE,
       PowerContactorEngaged := TRUE, JoystickOnline := TRUE, JoystickOperational := TRUE,
       HeartbeatIhmOk := TRUE, EncoderAvailable := TRUE, PhaseRotationOk := TRUE,
       TopPositionSensor := TRUE, FwdRevSpeedFeedbackOff := TRUE, BrakeFeedback := FALSE,
       JoystickYNeutral := TRUE, BenneHoldStillActive := FALSE, InReferencingMode := FALSE,
       CablePosM := 0.0, CfgCableLimitDescentM := -20.0, Homed := TRUE, TopLimitM := 8.5);
    ADVANCE_TIME(10000000);
    (* Scan 2 : surchauffe moteur (ThermalFeedback=TRUE) -> bit2 dans masque PowerCutOff *)
    fb(Enable := TRUE, Reset := FALSE, SyncEnable := FALSE,
       PowerContactorEngaged := TRUE, JoystickOnline := TRUE, JoystickOperational := TRUE,
       HeartbeatIhmOk := TRUE, EncoderAvailable := TRUE, PhaseRotationOk := TRUE,
       TopPositionSensor := TRUE, FwdRevSpeedFeedbackOff := TRUE, BrakeFeedback := FALSE,
       JoystickYNeutral := TRUE, BenneHoldStillActive := FALSE, InReferencingMode := FALSE,
       CablePosM := 0.0, CfgCableLimitDescentM := -20.0, Homed := TRUE, TopLimitM := 8.5,
       ThermalFeedback := TRUE);
    ASSERT_TRUE(fb.PowerCutOff, 'Surchauffe moteur (bit2) -> PowerCutOff (bit2 dans masque 16#2F84)');
    ASSERT_TRUE(fb.SafeStop, 'Surchauffe moteur -> SafeStop');
    (* Scan 3 : Reset acquitte *)
    ADVANCE_TIME(10000000);
    fb(Enable := TRUE, Reset := TRUE, SyncEnable := FALSE,
       PowerContactorEngaged := TRUE, JoystickOnline := TRUE, JoystickOperational := TRUE,
       HeartbeatIhmOk := TRUE, EncoderAvailable := TRUE, PhaseRotationOk := TRUE,
       TopPositionSensor := TRUE, FwdRevSpeedFeedbackOff := TRUE, BrakeFeedback := FALSE,
       JoystickYNeutral := TRUE, BenneHoldStillActive := FALSE, InReferencingMode := FALSE,
       CablePosM := 0.0, CfgCableLimitDescentM := -20.0, Homed := TRUE, TopLimitM := 8.5,
       ThermalFeedback := FALSE);
    ADVANCE_TIME(10000000);
    fb(Enable := TRUE, Reset := FALSE, SyncEnable := FALSE,
       PowerContactorEngaged := TRUE, JoystickOnline := TRUE, JoystickOperational := TRUE,
       HeartbeatIhmOk := TRUE, EncoderAvailable := TRUE, PhaseRotationOk := TRUE,
       TopPositionSensor := TRUE, FwdRevSpeedFeedbackOff := TRUE, BrakeFeedback := FALSE,
       JoystickYNeutral := TRUE, BenneHoldStillActive := FALSE, InReferencingMode := FALSE,
       CablePosM := 0.0, CfgCableLimitDescentM := -20.0, Homed := TRUE, TopLimitM := 8.5);
    ASSERT_FALSE(fb.Fault.Error, 'Reset acquitte la surchauffe');
    (* Scan 4 : sens oppose (bit14) -> SafeStop mais PAS PowerCutOff *)
    ADVANCE_TIME(10000000);
    fb(Enable := TRUE, Reset := FALSE, SyncEnable := FALSE,
       PowerContactorEngaged := TRUE, JoystickOnline := TRUE, JoystickOperational := TRUE,
       HeartbeatIhmOk := TRUE, EncoderAvailable := TRUE, PhaseRotationOk := TRUE,
       TopPositionSensor := TRUE, FwdRevSpeedFeedbackOff := TRUE, BrakeFeedback := FALSE,
       JoystickYNeutral := TRUE, BenneHoldStillActive := FALSE, InReferencingMode := FALSE,
       CablePosM := 0.0, CfgCableLimitDescentM := -20.0, Homed := TRUE, TopLimitM := 8.5,
       ReqAscent := TRUE, ReqDescend := FALSE, MovementCommanded := TRUE, MeasuredSpeedValid := TRUE,
       MeasuredSpeedSignedMps := -0.1);
    ADVANCE_TIME(500000000);
    fb(Enable := TRUE, Reset := FALSE, SyncEnable := FALSE,
       PowerContactorEngaged := TRUE, JoystickOnline := TRUE, JoystickOperational := TRUE,
       HeartbeatIhmOk := TRUE, EncoderAvailable := TRUE, PhaseRotationOk := TRUE,
       TopPositionSensor := TRUE, FwdRevSpeedFeedbackOff := TRUE, BrakeFeedback := FALSE,
       JoystickYNeutral := TRUE, BenneHoldStillActive := FALSE, InReferencingMode := FALSE,
       CablePosM := 0.0, CfgCableLimitDescentM := -20.0, Homed := TRUE, TopLimitM := 8.5,
       ReqAscent := TRUE, ReqDescend := FALSE, MovementCommanded := TRUE, MeasuredSpeedValid := TRUE,
       MeasuredSpeedSignedMps := -0.1);
    ASSERT_TRUE(fb.SafeStop, 'Sens oppose -> SafeStop');
    ASSERT_FALSE(fb.PowerCutOff, 'Sens oppose (bit14) -> PAS de PowerCutOff (hors masque 16#2F84)');
END_TEST

TEST 'TC-P10-010 SafeStop exclut bit3 (mou cable) si SyncEnable=FALSE'
    (* Scan 1 : regime nominal SyncEnable=FALSE *)
    fb(Enable := TRUE, Reset := FALSE, SyncEnable := FALSE,
       PowerContactorEngaged := TRUE, JoystickOnline := TRUE, JoystickOperational := TRUE,
       HeartbeatIhmOk := TRUE, EncoderAvailable := TRUE, PhaseRotationOk := TRUE,
       TopPositionSensor := TRUE, FwdRevSpeedFeedbackOff := TRUE, BrakeFeedback := FALSE,
       JoystickYNeutral := TRUE, BenneHoldStillActive := FALSE, InReferencingMode := FALSE,
       CablePosM := 0.0, CfgCableLimitDescentM := -20.0, Homed := TRUE, TopLimitM := 8.5);
    ADVANCE_TIME(10000000);
    (* Scan 2 : mou de cable (SlackCableDetected=TRUE), SyncEnable=FALSE -> bit3 exclu de SafeStop *)
    fb(Enable := TRUE, Reset := FALSE, SyncEnable := FALSE,
       PowerContactorEngaged := TRUE, JoystickOnline := TRUE, JoystickOperational := TRUE,
       HeartbeatIhmOk := TRUE, EncoderAvailable := TRUE, PhaseRotationOk := TRUE,
       TopPositionSensor := TRUE, FwdRevSpeedFeedbackOff := TRUE, BrakeFeedback := FALSE,
       JoystickYNeutral := TRUE, BenneHoldStillActive := FALSE, InReferencingMode := FALSE,
       CablePosM := 0.0, CfgCableLimitDescentM := -20.0, Homed := TRUE, TopLimitM := 8.5,
       SlackCableDetected := TRUE);
    ASSERT_FALSE(fb.SafeStop, 'Mou cable SyncEnable=FALSE -> PAS de SafeStop (bit3 exclu masque 16#FF97)');
    ASSERT_FALSE(fb.DescendPermit, 'Mou cable -> DescendPermit=FALSE (blocage descente)');
    ASSERT_TRUE(fb.AscentPermit, 'Mou cable -> AscentPermit reste TRUE');
    (* Scan 3 : cable retendu (SlackCableDetected=FALSE) -> blocage leve *)
    ADVANCE_TIME(10000000);
    fb(Enable := TRUE, Reset := FALSE, SyncEnable := FALSE,
       PowerContactorEngaged := TRUE, JoystickOnline := TRUE, JoystickOperational := TRUE,
       HeartbeatIhmOk := TRUE, EncoderAvailable := TRUE, PhaseRotationOk := TRUE,
       TopPositionSensor := TRUE, FwdRevSpeedFeedbackOff := TRUE, BrakeFeedback := FALSE,
       JoystickYNeutral := TRUE, BenneHoldStillActive := FALSE, InReferencingMode := FALSE,
       CablePosM := 0.0, CfgCableLimitDescentM := -20.0, Homed := TRUE, TopLimitM := 8.5,
       SlackCableDetected := FALSE);
    ASSERT_TRUE(fb.DescendPermit, 'Cable retendu -> DescendPermit=TRUE (blocage leve)');
END_TEST

TEST 'TC-P10-036.1 Warmup 3s : perte com operateur ignoree pendant 3s puis SafeStop'
    (* Scan 1 : Enable=TRUE, perte com operateur (JoystickOnline=FALSE) -> warmup en cours *)
    fb(Enable := TRUE, Reset := FALSE, SyncEnable := FALSE,
       PowerContactorEngaged := TRUE, JoystickOnline := FALSE, JoystickOperational := FALSE,
       HeartbeatIhmOk := FALSE, EncoderAvailable := TRUE, PhaseRotationOk := TRUE,
       TopPositionSensor := TRUE, FwdRevSpeedFeedbackOff := TRUE, BrakeFeedback := FALSE,
       JoystickYNeutral := TRUE, BenneHoldStillActive := FALSE, InReferencingMode := FALSE,
       CablePosM := 0.0, CfgCableLimitDescentM := -20.0, Homed := TRUE, TopLimitM := 8.5);
    ASSERT_FALSE(fb.SafeStop, 'Pendant warmup (<3s) : perte com ignoree -> pas de SafeStop');
    (* Scan 2 : 1s ecoulee, toujours < 3s *)
    ADVANCE_TIME(1000000000);
    fb(Enable := TRUE, Reset := FALSE, SyncEnable := FALSE,
       PowerContactorEngaged := TRUE, JoystickOnline := FALSE, JoystickOperational := FALSE,
       HeartbeatIhmOk := FALSE, EncoderAvailable := TRUE, PhaseRotationOk := TRUE,
       TopPositionSensor := TRUE, FwdRevSpeedFeedbackOff := TRUE, BrakeFeedback := FALSE,
       JoystickYNeutral := TRUE, BenneHoldStillActive := FALSE, InReferencingMode := FALSE,
       CablePosM := 0.0, CfgCableLimitDescentM := -20.0, Homed := TRUE, TopLimitM := 8.5);
    ASSERT_FALSE(fb.SafeStop, '1s : toujours pas de SafeStop');
    (* Scan 3 : apres 3s -> cause 0 active -> SafeStop *)
    ADVANCE_TIME(3000000000);
    fb(Enable := TRUE, Reset := FALSE, SyncEnable := FALSE,
       PowerContactorEngaged := TRUE, JoystickOnline := FALSE, JoystickOperational := FALSE,
       HeartbeatIhmOk := FALSE, EncoderAvailable := TRUE, PhaseRotationOk := TRUE,
       TopPositionSensor := TRUE, FwdRevSpeedFeedbackOff := TRUE, BrakeFeedback := FALSE,
       JoystickYNeutral := TRUE, BenneHoldStillActive := FALSE, InReferencingMode := FALSE,
       CablePosM := 0.0, CfgCableLimitDescentM := -20.0, Homed := TRUE, TopLimitM := 8.5);
    ASSERT_TRUE(fb.SafeStop, 'Apres 3s : perte com -> SafeStop');
    ASSERT_TRUE(fb.Fault.Error, 'Perte com -> Error');
END_TEST

TEST 'TC-P10-037.1 Gate Enable=FALSE : sorties forcees FALSE, latches preserves, re-Enable exige Reset'
    (* Scan 1 : regime nominal *)
    fb(Enable := TRUE, Reset := FALSE, SyncEnable := FALSE,
       PowerContactorEngaged := TRUE, JoystickOnline := TRUE, JoystickOperational := TRUE,
       HeartbeatIhmOk := TRUE, EncoderAvailable := TRUE, PhaseRotationOk := TRUE,
       TopPositionSensor := TRUE, FwdRevSpeedFeedbackOff := TRUE, BrakeFeedback := FALSE,
       JoystickYNeutral := TRUE, BenneHoldStillActive := FALSE, InReferencingMode := FALSE,
       CablePosM := 0.0, CfgCableLimitDescentM := -20.0, Homed := TRUE, TopLimitM := 8.5);
    ADVANCE_TIME(10000000);
    (* Scan 2 : declenche Meca A (derive >5.0m) - MES 2026-09-04 : seuil 2.0->5.0m *)
    fb(Enable := TRUE, Reset := FALSE, SyncEnable := FALSE,
       PowerContactorEngaged := TRUE, JoystickOnline := TRUE, JoystickOperational := TRUE,
       HeartbeatIhmOk := TRUE, EncoderAvailable := TRUE, PhaseRotationOk := TRUE,
       TopPositionSensor := TRUE, FwdRevSpeedFeedbackOff := TRUE, BrakeFeedback := FALSE,
       JoystickYNeutral := TRUE, BenneHoldStillActive := FALSE, InReferencingMode := FALSE,
       CablePosM := 6.0, CfgCableLimitDescentM := -20.0, Homed := TRUE, TopLimitM := 8.5);
    ASSERT_TRUE(fb.Fault.Error, 'Precondition : Meca A latchee');
    (* Scan 3 : Enable=FALSE -> sorties forcees FALSE, latch preserve *)
    ADVANCE_TIME(10000000);
    fb(Enable := FALSE, Reset := FALSE, SyncEnable := FALSE,
       PowerContactorEngaged := TRUE, JoystickOnline := TRUE, JoystickOperational := TRUE,
       HeartbeatIhmOk := TRUE, EncoderAvailable := TRUE, PhaseRotationOk := TRUE,
       TopPositionSensor := TRUE, FwdRevSpeedFeedbackOff := TRUE, BrakeFeedback := FALSE,
       JoystickYNeutral := TRUE, BenneHoldStillActive := FALSE, InReferencingMode := FALSE,
       CablePosM := 6.0, CfgCableLimitDescentM := -20.0, Homed := TRUE, TopLimitM := 8.5);
    ASSERT_FALSE(fb.SafeStop, 'Enable=FALSE -> SafeStop force FALSE');
    ASSERT_FALSE(fb.PowerCutOff, 'Enable=FALSE -> PowerCutOff force FALSE');
    ASSERT_FALSE(fb.Ready, 'Enable=FALSE -> Ready=FALSE');
    (* Scan 4 : re-Enable SANS Reset, cause disparue -> latch preserve (Ready=FALSE) *)
    ADVANCE_TIME(10000000);
    fb(Enable := TRUE, Reset := FALSE, SyncEnable := FALSE,
       PowerContactorEngaged := TRUE, JoystickOnline := TRUE, JoystickOperational := TRUE,
       HeartbeatIhmOk := TRUE, EncoderAvailable := TRUE, PhaseRotationOk := TRUE,
       TopPositionSensor := TRUE, FwdRevSpeedFeedbackOff := TRUE, BrakeFeedback := FALSE,
       JoystickYNeutral := TRUE, BenneHoldStillActive := FALSE, InReferencingMode := FALSE,
       CablePosM := 0.0, CfgCableLimitDescentM := -20.0, Homed := TRUE, TopLimitM := 8.5);
    ASSERT_FALSE(fb.Ready, 'Re-Enable sans Reset : latch preserve -> Ready=FALSE');
    ASSERT_TRUE(fb.Fault.Latched, 'Re-Enable sans Reset : defaut toujours latche');
    (* Scan 5 : front Reset -> acquitte *)
    ADVANCE_TIME(10000000);
    fb(Enable := TRUE, Reset := TRUE, SyncEnable := FALSE,
       PowerContactorEngaged := TRUE, JoystickOnline := TRUE, JoystickOperational := TRUE,
       HeartbeatIhmOk := TRUE, EncoderAvailable := TRUE, PhaseRotationOk := TRUE,
       TopPositionSensor := TRUE, FwdRevSpeedFeedbackOff := TRUE, BrakeFeedback := FALSE,
       JoystickYNeutral := TRUE, BenneHoldStillActive := FALSE, InReferencingMode := FALSE,
       CablePosM := 0.0, CfgCableLimitDescentM := -20.0, Homed := TRUE, TopLimitM := 8.5);
    ADVANCE_TIME(10000000);
    fb(Enable := TRUE, Reset := FALSE, SyncEnable := FALSE,
       PowerContactorEngaged := TRUE, JoystickOnline := TRUE, JoystickOperational := TRUE,
       HeartbeatIhmOk := TRUE, EncoderAvailable := TRUE, PhaseRotationOk := TRUE,
       TopPositionSensor := TRUE, FwdRevSpeedFeedbackOff := TRUE, BrakeFeedback := FALSE,
       JoystickYNeutral := TRUE, BenneHoldStillActive := FALSE, InReferencingMode := FALSE,
       CablePosM := 0.0, CfgCableLimitDescentM := -20.0, Homed := TRUE, TopLimitM := 8.5);
    ASSERT_TRUE(fb.Ready, 'Reset front -> Ready=TRUE');
    ASSERT_FALSE(fb.Fault.Error, 'Reset front -> plus d erreur');
END_TEST

TEST 'TC-P10-044.1 Mou cable : SyncEnable=FALSE -> DescendPermit=FALSE, AscentPermit autorise, blocage leve au retension'
    (* Scan 1 : regime nominal SyncEnable=FALSE *)
    fb(Enable := TRUE, Reset := FALSE, SyncEnable := FALSE,
       PowerContactorEngaged := TRUE, JoystickOnline := TRUE, JoystickOperational := TRUE,
       HeartbeatIhmOk := TRUE, EncoderAvailable := TRUE, PhaseRotationOk := TRUE,
       TopPositionSensor := TRUE, FwdRevSpeedFeedbackOff := TRUE, BrakeFeedback := FALSE,
       JoystickYNeutral := TRUE, BenneHoldStillActive := FALSE, InReferencingMode := FALSE,
       CablePosM := 0.0, CfgCableLimitDescentM := -20.0, Homed := TRUE, TopLimitM := 8.5);
    ADVANCE_TIME(10000000);
    (* Scan 2 : mou de cable -> blocage descente, montee autorisee *)
    fb(Enable := TRUE, Reset := FALSE, SyncEnable := FALSE,
       PowerContactorEngaged := TRUE, JoystickOnline := TRUE, JoystickOperational := TRUE,
       HeartbeatIhmOk := TRUE, EncoderAvailable := TRUE, PhaseRotationOk := TRUE,
       TopPositionSensor := TRUE, FwdRevSpeedFeedbackOff := TRUE, BrakeFeedback := FALSE,
       JoystickYNeutral := TRUE, BenneHoldStillActive := FALSE, InReferencingMode := FALSE,
       CablePosM := 0.0, CfgCableLimitDescentM := -20.0, Homed := TRUE, TopLimitM := 8.5,
       SlackCableDetected := TRUE);
    ASSERT_FALSE(fb.DescendPermit, 'Mou cable -> DescendPermit=FALSE');
    ASSERT_TRUE(fb.AscentPermit, 'Mou cable -> AscentPermit=TRUE (montee autorisee)');
    ASSERT_FALSE(fb.SafeStop, 'Mou cable SyncEnable=FALSE -> pas de SafeStop (bit3 exclu)');
    (* Scan 3 : cable retendu (M2_TensionedCable_DI=TRUE) -> blocage leve *)
    ADVANCE_TIME(10000000);
    fb(Enable := TRUE, Reset := FALSE, SyncEnable := FALSE,
       PowerContactorEngaged := TRUE, JoystickOnline := TRUE, JoystickOperational := TRUE,
       HeartbeatIhmOk := TRUE, EncoderAvailable := TRUE, PhaseRotationOk := TRUE,
       TopPositionSensor := TRUE, FwdRevSpeedFeedbackOff := TRUE, BrakeFeedback := FALSE,
       JoystickYNeutral := TRUE, BenneHoldStillActive := FALSE, InReferencingMode := FALSE,
       CablePosM := 0.0, CfgCableLimitDescentM := -20.0, Homed := TRUE, TopLimitM := 8.5,
       SlackCableDetected := FALSE);
    ASSERT_TRUE(fb.DescendPermit, 'Cable retendu -> DescendPermit=TRUE');
END_TEST

TEST 'TC-P10-051.1 Chaine PowerCutOff bout-en-bout : FB produit la coupure, chaine PRG_04->PRG_06->AU = essai site'
    (* (essai site — stub) : la preuve bout-en-bout (demande PRG_04 -> agregation PRG_06 -> coupure AU)
       n est pas automatisable en boite noire FB. On verifie ici la brique amont : le FB produit
       bien PowerCutOff sur une cause du masque 16#2F84, condition necessaire de la chaine. *)
    fb(Enable := TRUE, Reset := FALSE, SyncEnable := FALSE,
       PowerContactorEngaged := TRUE, JoystickOnline := TRUE, JoystickOperational := TRUE,
       HeartbeatIhmOk := TRUE, EncoderAvailable := TRUE, PhaseRotationOk := TRUE,
       TopPositionSensor := TRUE, FwdRevSpeedFeedbackOff := TRUE, BrakeFeedback := FALSE,
       JoystickYNeutral := TRUE, BenneHoldStillActive := FALSE, InReferencingMode := FALSE,
       CablePosM := 0.0, CfgCableLimitDescentM := -20.0, Homed := TRUE, TopLimitM := 8.5);
    ADVANCE_TIME(10000000);
    fb(Enable := TRUE, Reset := FALSE, SyncEnable := FALSE,
       PowerContactorEngaged := TRUE, JoystickOnline := TRUE, JoystickOperational := TRUE,
       HeartbeatIhmOk := TRUE, EncoderAvailable := TRUE, PhaseRotationOk := TRUE,
       TopPositionSensor := TRUE, FwdRevSpeedFeedbackOff := TRUE, BrakeFeedback := FALSE,
       JoystickYNeutral := TRUE, BenneHoldStillActive := FALSE, InReferencingMode := FALSE,
       CablePosM := 6.0, CfgCableLimitDescentM := -20.0, Homed := TRUE, TopLimitM := 8.5);
    ASSERT_TRUE(fb.PowerCutOff, 'Cause masque 16#2F84 -> PowerCutOff produit (brique amont de la chaine)');
    ASSERT_TRUE(fb.SafeStop, 'Cause masque -> SafeStop');
END_TEST

TEST 'TC-P10-052 Limite legale : BypassProcess simu ne leve pas le verrou sous -15m'
    (* Regression T197 : SimulationBypassActive arme BypassProcess pour eviter les
       faux defauts mecaniques du banc. Ce bypass de groupe ne doit pas neutraliser
       la limite legale; seul BypassLimitLegal est habilite a le faire. *)
    fb(Enable := TRUE, Reset := FALSE, SyncEnable := TRUE,
       PowerContactorEngaged := TRUE, JoystickOnline := TRUE, JoystickOperational := TRUE,
       HeartbeatIhmOk := TRUE, EncoderAvailable := TRUE, PhaseRotationOk := TRUE,
       TopPositionSensor := TRUE, FwdRevSpeedFeedbackOff := TRUE, BrakeFeedback := FALSE,
       JoystickYNeutral := TRUE, BenneHoldStillActive := FALSE, BenneBusy := FALSE,
       OtherWinchInhibited := FALSE, InReferencingMode := FALSE,
       CablePosM := -15.1, CfgCableLimitDescentM := -20.0,
       LimitLegalReached := TRUE, Homed := TRUE, TopLimitM := 8.5,
       BypassProcess := TRUE, BypassLimitLegal := FALSE);
    ADVANCE_TIME(10000000);
    fb(Enable := TRUE, Reset := FALSE, SyncEnable := TRUE,
       PowerContactorEngaged := TRUE, JoystickOnline := TRUE, JoystickOperational := TRUE,
       HeartbeatIhmOk := TRUE, EncoderAvailable := TRUE, PhaseRotationOk := TRUE,
       TopPositionSensor := TRUE, FwdRevSpeedFeedbackOff := TRUE, BrakeFeedback := FALSE,
       JoystickYNeutral := TRUE, BenneHoldStillActive := FALSE, BenneBusy := FALSE,
       OtherWinchInhibited := FALSE, InReferencingMode := FALSE,
       CablePosM := -15.1, CfgCableLimitDescentM := -20.0,
       LimitLegalReached := TRUE, Homed := TRUE, TopLimitM := 8.5,
       BypassProcess := TRUE, BypassLimitLegal := FALSE);
    ASSERT_FALSE(fb.DescendPermit, 'BypassProcess seul ne doit pas autoriser la descente sous la limite legale');
END_TEST

TEST 'TC-P10-053 Limite legale : bypass dedie explicite autorise uniquement le test MAINT_N2'
    (* Le bypass legal dedie conserve le comportement de mise en service; il est
       gate par MAINT_N2 dans PRG_04 avant d arriver ici. *)
    fb(Enable := TRUE, Reset := FALSE, SyncEnable := TRUE,
       PowerContactorEngaged := TRUE, JoystickOnline := TRUE, JoystickOperational := TRUE,
       HeartbeatIhmOk := TRUE, EncoderAvailable := TRUE, PhaseRotationOk := TRUE,
       TopPositionSensor := TRUE, FwdRevSpeedFeedbackOff := TRUE, BrakeFeedback := FALSE,
       JoystickYNeutral := TRUE, BenneHoldStillActive := FALSE, BenneBusy := FALSE,
       OtherWinchInhibited := FALSE, InReferencingMode := FALSE,
       CablePosM := -15.1, CfgCableLimitDescentM := -20.0,
       LimitLegalReached := TRUE, Homed := TRUE, TopLimitM := 8.5,
       BypassProcess := TRUE, BypassLimitLegal := TRUE);
    ADVANCE_TIME(10000000);
    fb(Enable := TRUE, Reset := FALSE, SyncEnable := TRUE,
       PowerContactorEngaged := TRUE, JoystickOnline := TRUE, JoystickOperational := TRUE,
       HeartbeatIhmOk := TRUE, EncoderAvailable := TRUE, PhaseRotationOk := TRUE,
       TopPositionSensor := TRUE, FwdRevSpeedFeedbackOff := TRUE, BrakeFeedback := FALSE,
       JoystickYNeutral := TRUE, BenneHoldStillActive := FALSE, BenneBusy := FALSE,
       OtherWinchInhibited := FALSE, InReferencingMode := FALSE,
       CablePosM := -15.1, CfgCableLimitDescentM := -20.0,
       LimitLegalReached := TRUE, Homed := TRUE, TopLimitM := 8.5,
       BypassProcess := TRUE, BypassLimitLegal := TRUE);
    ASSERT_TRUE(fb.DescendPermit, 'BypassLimitLegal explicite autorise le test de descente');
END_TEST

TEST 'T387-001 Meca B mode boutons MAINT_N2 : commande bouton (joystick neutre) -> PAS de faux arrêt non confirmé'
    (* T387 - Repro faux positif : commande PAR BOUTON IHM. Le joystick reste au
       neutre (JoystickYNeutral=TRUE) pendant que la commande de mouvement est
       active (MovementCommanded=TRUE, ReqAscent=TRUE, contacteurs engages +
       frein ouvert, vitesse valide vers le haut). MecaB ne doit PAS se
       declencher : le treuil est commande (avant fix T387 : MecaB latche = ROUGE). *)
    (* RAZ des latches partages venant des tests precedents (instance fb unique) *)
    fb(Enable := TRUE, Reset := TRUE, SyncEnable := FALSE,
       PowerContactorEngaged := TRUE, JoystickOnline := TRUE, JoystickOperational := TRUE,
       HeartbeatIhmOk := TRUE, EncoderAvailable := TRUE, PhaseRotationOk := TRUE,
       TopPositionSensor := FALSE, FwdRevSpeedFeedbackOff := TRUE, BrakeFeedback := FALSE,
       JoystickYNeutral := TRUE, BenneHoldStillActive := FALSE, InReferencingMode := FALSE,
       CablePosM := 0.0, CfgCableLimitDescentM := -20.0, Homed := TRUE, TopLimitM := 8.5);
    ADVANCE_TIME(10000000);
    (* Scan nominal reference *)
    fb(Enable := TRUE, Reset := FALSE, SyncEnable := FALSE,
       PowerContactorEngaged := TRUE, JoystickOnline := TRUE, JoystickOperational := TRUE,
       HeartbeatIhmOk := TRUE, EncoderAvailable := TRUE, PhaseRotationOk := TRUE,
       TopPositionSensor := FALSE, FwdRevSpeedFeedbackOff := TRUE, BrakeFeedback := FALSE,
       JoystickYNeutral := TRUE, BenneHoldStillActive := FALSE, InReferencingMode := FALSE,
       CablePosM := 0.0, CfgCableLimitDescentM := -20.0, Homed := TRUE, TopLimitM := 8.5);
    ADVANCE_TIME(3000000000);
    (* Commande bouton active : joystick neutre (boutons) + mouvement commande *)
    fb(Enable := TRUE, Reset := FALSE, SyncEnable := FALSE,
       PowerContactorEngaged := TRUE, JoystickOnline := TRUE, JoystickOperational := TRUE,
       HeartbeatIhmOk := TRUE, EncoderAvailable := TRUE, PhaseRotationOk := TRUE,
       TopPositionSensor := FALSE, FwdRevSpeedFeedbackOff := FALSE, BrakeFeedback := TRUE,
       JoystickYNeutral := TRUE, BenneHoldStillActive := FALSE, InReferencingMode := FALSE,
       CablePosM := 0.0, CfgCableLimitDescentM := -20.0, Homed := TRUE, TopLimitM := 8.5,
       MeasuredSpeedValid := TRUE, MeasuredSpeedMps := 0.5, MeasuredSpeedSignedMps := 0.5,
       ReqAscent := TRUE, ReqDescend := FALSE, MovementCommanded := TRUE);
    ADVANCE_TIME(3000000000);
    fb(Enable := TRUE, Reset := FALSE, SyncEnable := FALSE,
       PowerContactorEngaged := TRUE, JoystickOnline := TRUE, JoystickOperational := TRUE,
       HeartbeatIhmOk := TRUE, EncoderAvailable := TRUE, PhaseRotationOk := TRUE,
       TopPositionSensor := FALSE, FwdRevSpeedFeedbackOff := FALSE, BrakeFeedback := TRUE,
       JoystickYNeutral := TRUE, BenneHoldStillActive := FALSE, InReferencingMode := FALSE,
       CablePosM := 0.0, CfgCableLimitDescentM := -20.0, Homed := TRUE, TopLimitM := 8.5,
       MeasuredSpeedValid := TRUE, MeasuredSpeedMps := 0.5, MeasuredSpeedSignedMps := 0.5,
       ReqAscent := TRUE, ReqDescend := FALSE, MovementCommanded := TRUE);
    ASSERT_TRUE(fb.MecaBElapsedTime < T#3s, 'Mode boutons MAINT_N2 (commande bouton) : MecaB ne doit PAS armer -> MecaBElapsedTime < 3s. ROUGE avant fix / VERT apres (T387).');
    ASSERT_FALSE((fb.Fault.LatchedId AND 16#0100) <> 0, 'Mode boutons MAINT_N2 : pas de cause MecaB (bit 0x100) pendant commande bouton');
END_TEST

TEST 'T387-FB-002 Grant fenetre benne : BucketCloseAscentGrant relaxe ETROITEMENT la butee haute MATERIELLE M2'
    (* T387 Fenetre benne (AC1/AC2) : fermer la benne = M2 monte relatif a M1 FIXE -> l'ensemble M1/M2
       ne change PAS d'altitude, donc en position haute la butee materielle M2 ne doit PAS bloquer la
       fermeture sur place. Le grant (calcule dans PRG_04 sous 4 verrous) est cable TRUE uniquement
       sur l'instance M2 et FALSE sur M1 (AC3 : le FdC materiel haut M1 reste la barriere absolue).
       Boite noire FB : grant=TRUE -> AscentPermit relaxe ; grant=FALSE -> barriere active.
       ⛔ ROUGE avant fix (AscentPermit ignore encore le grant) / VERT apres. *)
    (* RAZ latches de l'instance partagee. *)
    fb(Enable := TRUE, Reset := TRUE, SyncEnable := FALSE,
       PowerContactorEngaged := TRUE, JoystickOnline := TRUE, JoystickOperational := TRUE,
       HeartbeatIhmOk := TRUE, EncoderAvailable := TRUE, PhaseRotationOk := TRUE,
       TopPositionSensor := FALSE, FwdRevSpeedFeedbackOff := TRUE, BrakeFeedback := FALSE,
       JoystickYNeutral := TRUE, BenneHoldStillActive := FALSE, InReferencingMode := FALSE,
       CablePosM := 0.0, CfgCableLimitDescentM := -20.0, Homed := TRUE, TopLimitM := 8.5,
       BucketCloseAscentGrant := FALSE);
    ADVANCE_TIME(10000000);
    (* Capture : FdC haut atteint + grant=FALSE -> barriere active. *)
    fb(Enable := TRUE, Reset := FALSE, SyncEnable := FALSE,
       PowerContactorEngaged := TRUE, JoystickOnline := TRUE, JoystickOperational := TRUE,
       HeartbeatIhmOk := TRUE, EncoderAvailable := TRUE, PhaseRotationOk := TRUE,
       TopPositionSensor := FALSE, FwdRevSpeedFeedbackOff := TRUE, BrakeFeedback := FALSE,
       JoystickYNeutral := TRUE, BenneHoldStillActive := FALSE, InReferencingMode := FALSE,
       CablePosM := 0.0, CfgCableLimitDescentM := -20.0, Homed := TRUE, TopLimitM := 8.5,
       BucketCloseAscentGrant := FALSE);
    ASSERT_FALSE(fb.AscentPermit, 'FdC haut atteint + grant=FALSE -> AscentPermit FALSE (barriere active)');
    (* Scan : grant=TRUE (fenetre benne active) -> barriere MATERIELLE relaxee ETROITEMENT. *)
    ADVANCE_TIME(10000000);
    fb(Enable := TRUE, Reset := FALSE, SyncEnable := FALSE,
       PowerContactorEngaged := TRUE, JoystickOnline := TRUE, JoystickOperational := TRUE,
       HeartbeatIhmOk := TRUE, EncoderAvailable := TRUE, PhaseRotationOk := TRUE,
       TopPositionSensor := FALSE, FwdRevSpeedFeedbackOff := TRUE, BrakeFeedback := FALSE,
       JoystickYNeutral := TRUE, BenneHoldStillActive := FALSE, InReferencingMode := FALSE,
       CablePosM := 0.0, CfgCableLimitDescentM := -20.0, Homed := TRUE, TopLimitM := 8.5,
       BucketCloseAscentGrant := TRUE);
    ASSERT_TRUE(fb.AscentPermit, 'Fenetre benne grant=TRUE -> AscentPermit relaxe malgre le FdC haut (M2, AC2)');
    // Le grant ne BYPASSE pas la cause : le FdC haut (cause 5, bit 16#0020) reste VIVANT et
    // informe (seul le PERMIS est relaxe). Erreur live bit5 attendue -> jamais un bypass total.
    ASSERT_TRUE((fb.Fault.ErrorId AND 16#0020) <> 0, 'Fenetre benne : cause 5 (FdC haut) reste vive (grant relaxe le permis, pas la cause)');
    ASSERT_FALSE(fb.Fault.Latched, 'Fenetre benne : cause live non latchable (Latching=FALSE) -> aucun defaut a acquitter');
    (* Scan : retour grant=FALSE (hors fenetre) -> la barriere reprend immediatement. *)
    ADVANCE_TIME(10000000);
    fb(Enable := TRUE, Reset := FALSE, SyncEnable := FALSE,
       PowerContactorEngaged := TRUE, JoystickOnline := TRUE, JoystickOperational := TRUE,
       HeartbeatIhmOk := TRUE, EncoderAvailable := TRUE, PhaseRotationOk := TRUE,
       TopPositionSensor := FALSE, FwdRevSpeedFeedbackOff := TRUE, BrakeFeedback := FALSE,
       JoystickYNeutral := TRUE, BenneHoldStillActive := FALSE, InReferencingMode := FALSE,
       CablePosM := 0.0, CfgCableLimitDescentM := -20.0, Homed := TRUE, TopLimitM := 8.5,
       BucketCloseAscentGrant := FALSE);
    ASSERT_FALSE(fb.AscentPermit, 'grant=FALSE (hors fenetre) -> barriere M2 active immediatement (AC2 bornee)');
END_TEST

(* ---- FB_SpeedStep_test.st ---- *)
(* =======================================================================
   test_fb_speedstep.st — T181-07 : bornes Min/Max du décodeur palier
   ======================================================================= *)

SETUP
VAR
    fb : FB_SpeedStep;
    Table : ST_SpeedStepTable;
END_VAR
END_SETUP

TEST 'TC-P10-T181-07a Defaut retro-compatible : demande 4 -> palier 4'
    Table.StepThreshold_Pct[1] := 10.0;
    Table.StepThreshold_Pct[2] := 30.0;
    Table.StepThreshold_Pct[3] := 50.0;
    Table.StepThreshold_Pct[4] := 70.0;
    Table.StepThreshold_Pct[5] := 90.0;
    Table.P4R1 := TRUE;

    fb(Enable := TRUE, SpeedStepReq := 4, Table := Table, MaxStepNumber := 5);
    ASSERT_EQ(fb.StepNumber, 4, 'Defaut Min=1 : demande 4 conservee');
    ASSERT_TRUE(fb.Contactor1, 'Table palier 4 lue');
END_TEST

TEST 'TC-P10-T181-07b Precedence plafond : plancher 3 + plafond 1 -> palier 1'
    Table.StepThreshold_Pct[1] := 10.0;
    Table.StepThreshold_Pct[2] := 30.0;
    Table.StepThreshold_Pct[3] := 50.0;
    Table.StepThreshold_Pct[4] := 70.0;
    Table.StepThreshold_Pct[5] := 90.0;
    Table.P1R1 := TRUE;

    fb(Enable := TRUE, SpeedStepReq := 5, Table := Table, MinStepNumber := 3, MaxStepNumber := 1);
    ASSERT_EQ(fb.StepNumber, 1, 'Le plafond securite gagne sur le plancher');
    ASSERT_TRUE(fb.Contactor1, 'Table palier 1 lue');
END_TEST

TEST 'TC-P10-T181-07c Relache : Enable FALSE force le palier 0'
    Table.StepThreshold_Pct[1] := 10.0;
    Table.StepThreshold_Pct[2] := 30.0;
    Table.StepThreshold_Pct[3] := 50.0;
    Table.StepThreshold_Pct[4] := 70.0;
    Table.StepThreshold_Pct[5] := 90.0;
    Table.P3R1 := TRUE;

    fb(Enable := FALSE, SpeedStepReq := 5, Table := Table, MinStepNumber := 3, MaxStepNumber := 5);
    ASSERT_EQ(fb.StepNumber, 0, 'Relache : le plancher ne maintient aucun palier');
    ASSERT_FALSE(fb.Contactor1, 'Relache : contacteur 1 coupe');
END_TEST

TEST 'TC-P10-T181-07d Bornes : requete hors plage reste dans 0..5'
    Table.StepThreshold_Pct[1] := 10.0;
    Table.StepThreshold_Pct[2] := 30.0;
    Table.StepThreshold_Pct[3] := 50.0;
    Table.StepThreshold_Pct[4] := 70.0;
    Table.StepThreshold_Pct[5] := 90.0;
    Table.P5R1 := TRUE;

    fb(Enable := TRUE, SpeedStepReq := 99, Table := Table, MinStepNumber := -3, MaxStepNumber := 99);
    ASSERT_EQ(fb.StepNumber, 5, 'Requete et plafond hauts bornes a 5');
    fb(Enable := TRUE, SpeedStepReq := -1, Table := Table, MinStepNumber := 5, MaxStepNumber := 5);
    ASSERT_EQ(fb.StepNumber, 0, 'Requete nulle ou negative reste a 0');
END_TEST

(* ---- FB_SyncContactor_test.st ---- *)
SETUP
VAR
    fb : FB_SyncContactor;
END_VAR
END_SETUP

TEST 'TC-P10-SYNC-01 Discordance Niveau 1 SafeStop'
    (* Etape 0 : Regime symetrique P2 monte *)
    fb(Enable := TRUE, Reset := FALSE, SyncEnable := TRUE,
       RelayFwdM1 := TRUE, RelayFwdM2 := TRUE,
       RelayRevM1 := FALSE, RelayRevM2 := FALSE,
       Contactor1_M1 := TRUE, Contactor1_M2 := TRUE,
       Contactor2_M1 := FALSE, Contactor2_M2 := FALSE,
       Contactor3_M1 := FALSE, Contactor3_M2 := FALSE,
       Contactor4_M1 := FALSE, Contactor4_M2 := FALSE,
       BypassGlobal := FALSE);
    ASSERT_FALSE(fb.ContactorMismatch, 'Regime symetrique -> pas de discordance');
    ASSERT_EQ(fb.Diag.MismatchLevel, 0, 'MismatchLevel = 0');

    (* Etape 1 : Apparition discordance M1 passe P3 (K2) *)
    ADVANCE_TIME(10000000);
    fb(Enable := TRUE, Reset := FALSE, SyncEnable := TRUE,
       RelayFwdM1 := TRUE, RelayFwdM2 := TRUE,
       RelayRevM1 := FALSE, RelayRevM2 := FALSE,
       Contactor1_M1 := TRUE, Contactor1_M2 := TRUE,
       Contactor2_M1 := TRUE, Contactor2_M2 := FALSE,
       Contactor3_M1 := FALSE, Contactor3_M2 := FALSE,
       Contactor4_M1 := FALSE, Contactor4_M2 := FALSE,
       BypassGlobal := FALSE);
    ASSERT_TRUE(fb.Diag.Step2Mismatch, 'Step2Mismatch detecte');

    (* Etape 2 : Filtrage debounce avant 500ms *)
    ADVANCE_TIME(250000000);
    fb(Enable := TRUE, Reset := FALSE, SyncEnable := TRUE,
       RelayFwdM1 := TRUE, RelayFwdM2 := TRUE,
       RelayRevM1 := FALSE, RelayRevM2 := FALSE,
       Contactor1_M1 := TRUE, Contactor1_M2 := TRUE,
       Contactor2_M1 := TRUE, Contactor2_M2 := FALSE,
       Contactor3_M1 := FALSE, Contactor3_M2 := FALSE,
       Contactor4_M1 := FALSE, Contactor4_M2 := FALSE,
       BypassGlobal := FALSE);
    ASSERT_FALSE(fb.ContactorMismatch, 'Pas de SafeStop avant debounce 500ms');

    (* Etape 3 : Declenchement SafeStop apres 500ms *)
    ADVANCE_TIME(260000000);
    fb(Enable := TRUE, Reset := FALSE, SyncEnable := TRUE,
       RelayFwdM1 := TRUE, RelayFwdM2 := TRUE,
       RelayRevM1 := FALSE, RelayRevM2 := FALSE,
       Contactor1_M1 := TRUE, Contactor1_M2 := TRUE,
       Contactor2_M1 := TRUE, Contactor2_M2 := FALSE,
       Contactor3_M1 := FALSE, Contactor3_M2 := FALSE,
       Contactor4_M1 := FALSE, Contactor4_M2 := FALSE,
       BypassGlobal := FALSE);
    ASSERT_TRUE(fb.ContactorMismatch, 'ContactorMismatch=TRUE apres 500ms');
    ASSERT_FALSE(fb.ContactorMismatchEscalated, 'Pas encore escalade');
    ASSERT_EQ(fb.Diag.MismatchLevel, 1, 'MismatchLevel = 1 (SafeStop)');
END_TEST

TEST 'TC-P10-SYNC-02 Escalade Niveau 2 PowerCutOff'
    (* Etablissement Niveau 1 *)
    fb(Enable := TRUE, Reset := FALSE, SyncEnable := TRUE,
       RelayFwdM1 := TRUE, RelayFwdM2 := TRUE,
       RelayRevM1 := FALSE, RelayRevM2 := FALSE,
       Contactor1_M1 := TRUE, Contactor1_M2 := FALSE,
       Contactor2_M1 := FALSE, Contactor2_M2 := FALSE,
       Contactor3_M1 := FALSE, Contactor3_M2 := FALSE,
       Contactor4_M1 := FALSE, Contactor4_M2 := FALSE,
       BypassGlobal := FALSE);
    ADVANCE_TIME(550000000);
    fb(Enable := TRUE, Reset := FALSE, SyncEnable := TRUE,
       RelayFwdM1 := TRUE, RelayFwdM2 := TRUE,
       RelayRevM1 := FALSE, RelayRevM2 := FALSE,
       Contactor1_M1 := TRUE, Contactor1_M2 := FALSE,
       Contactor2_M1 := FALSE, Contactor2_M2 := FALSE,
       Contactor3_M1 := FALSE, Contactor3_M2 := FALSE,
       Contactor4_M1 := FALSE, Contactor4_M2 := FALSE,
       BypassGlobal := FALSE);
    ASSERT_TRUE(fb.ContactorMismatch, 'Niveau 1 etabli');

    (* Persistance pendant 3s supplementaires -> Escalade *)
    ADVANCE_TIME(3050000000);
    fb(Enable := TRUE, Reset := FALSE, SyncEnable := TRUE,
       RelayFwdM1 := TRUE, RelayFwdM2 := TRUE,
       RelayRevM1 := FALSE, RelayRevM2 := FALSE,
       Contactor1_M1 := TRUE, Contactor1_M2 := FALSE,
       Contactor2_M1 := FALSE, Contactor2_M2 := FALSE,
       Contactor3_M1 := FALSE, Contactor3_M2 := FALSE,
       Contactor4_M1 := FALSE, Contactor4_M2 := FALSE,
       BypassGlobal := FALSE);
    ASSERT_TRUE(fb.ContactorMismatchEscalated, 'ContactorMismatchEscalated=TRUE apres 3s');
    ASSERT_EQ(fb.Diag.MismatchLevel, 2, 'MismatchLevel = 2 (PowerCutOff)');
END_TEST

TEST 'TC-P10-SYNC-03 Jog unitaire Inhibition'
    (* Jog M1 seul : M2 non commande et SyncEnable=FALSE *)
    fb(Enable := TRUE, Reset := FALSE, SyncEnable := FALSE,
       RelayFwdM1 := TRUE, RelayFwdM2 := FALSE,
       RelayRevM1 := FALSE, RelayRevM2 := FALSE,
       Contactor1_M1 := TRUE, Contactor1_M2 := FALSE,
       Contactor2_M1 := FALSE, Contactor2_M2 := FALSE,
       Contactor3_M1 := FALSE, Contactor3_M2 := FALSE,
       Contactor4_M1 := FALSE, Contactor4_M2 := FALSE,
       BypassGlobal := FALSE);
    ADVANCE_TIME(1000000000);
    fb(Enable := TRUE, Reset := FALSE, SyncEnable := FALSE,
       RelayFwdM1 := TRUE, RelayFwdM2 := FALSE,
       RelayRevM1 := FALSE, RelayRevM2 := FALSE,
       Contactor1_M1 := TRUE, Contactor1_M2 := FALSE,
       Contactor2_M1 := FALSE, Contactor2_M2 := FALSE,
       Contactor3_M1 := FALSE, Contactor3_M2 := FALSE,
       Contactor4_M1 := FALSE, Contactor4_M2 := FALSE,
       BypassGlobal := FALSE);
    ASSERT_FALSE(fb.ContactorMismatch, 'Jog unitaire M1 -> Surveillance neutralisee');
    ASSERT_EQ(fb.Diag.MismatchLevel, 0, 'MismatchLevel = 0');
END_TEST

TEST 'TC-P10-SYNC-04 Bypass Global'
    fb(Enable := TRUE, Reset := FALSE, SyncEnable := TRUE,
       RelayFwdM1 := TRUE, RelayFwdM2 := FALSE,
       RelayRevM1 := FALSE, RelayRevM2 := TRUE,
       Contactor1_M1 := TRUE, Contactor1_M2 := FALSE,
       Contactor2_M1 := TRUE, Contactor2_M2 := FALSE,
       Contactor3_M1 := TRUE, Contactor3_M2 := FALSE,
       Contactor4_M1 := TRUE, Contactor4_M2 := FALSE,
       BypassGlobal := TRUE);
    ADVANCE_TIME(5000000000);
    fb(Enable := TRUE, Reset := FALSE, SyncEnable := TRUE,
       RelayFwdM1 := TRUE, RelayFwdM2 := FALSE,
       RelayRevM1 := FALSE, RelayRevM2 := TRUE,
       Contactor1_M1 := TRUE, Contactor1_M2 := FALSE,
       Contactor2_M1 := TRUE, Contactor2_M2 := FALSE,
       Contactor3_M1 := TRUE, Contactor3_M2 := FALSE,
       Contactor4_M1 := TRUE, Contactor4_M2 := FALSE,
       BypassGlobal := TRUE);
    ASSERT_FALSE(fb.ContactorMismatch, 'BypassGlobal -> Pas de mismatch');
    ASSERT_FALSE(fb.ContactorMismatchEscalated, 'BypassGlobal -> Pas d escalade');
    ASSERT_EQ(fb.Diag.MismatchLevel, 0, 'MismatchLevel = 0');
END_TEST

(* ---- FB_Winch_Symmetry_test.st ---- *)
(* =======================================================================
   test_fb_winch_symmetry.st -- T181-18 D11 : macro TC FB_Winch_Symmetry (F10.06)
   Observateur passif de symetrie / synchronisme M1-M2. Aucune action securite.
   Qualification : commande stable des 2 treuils, meme sens, au-dela de
   MinimumCommandTime_Ms (defaut 1000 ms) et vitesse au-dessus de MinimumSpeed_Mps.
   Les ecarts sont calcules a l arret.
   ======================================================================= *)

SETUP
VAR
    fb  : FB_Winch_Symmetry;
    Cfg : ST_fbWinch_Symmetry_Cfg;
    Dat : ST_fbWinch_Symmetry_Data;
END_VAR
END_SETUP

TEST 'TC-P10-T181-18a Cycle symetrique -> SymmetryValid et SymmetryOk'
    Cfg.MinimumCommandTime_Ms := 300;
    Cfg.MinimumSpeed_Mps := 0.05;
    Cfg.DeltaStartDelay_Ms := 100; Cfg.DeltaBrakeReleaseTime_Ms := 100;
    Cfg.DeltaBrakeApplyTime_Ms := 100; Cfg.DeltaStopDistance_Mm := 100;
    Cfg.DeltaStopTime_Ms := 200;
    fb(Reset := TRUE, M1CommandActive := FALSE, M2CommandActive := FALSE, M1Direction := 0, M2Direction := 0,
       M1BrakeCmd := FALSE, M2BrakeCmd := FALSE, M1BrakeApplied := TRUE, M2BrakeApplied := TRUE,
       M1Position_M := 0.0, M2Position_M := 0.0, M1Speed_Mps := 0.0, M2Speed_Mps := 0.0,
       SyncDeviation_M := 0.0, Config := Cfg, Data := Dat);
    fb(Reset := FALSE, M1CommandActive := TRUE, M2CommandActive := TRUE, M1Direction := 1, M2Direction := 1,
       M1BrakeCmd := TRUE, M2BrakeCmd := TRUE, M1BrakeApplied := FALSE, M2BrakeApplied := FALSE,
       M1Position_M := 0.0, M2Position_M := 0.0, M1Speed_Mps := 1.0, M2Speed_Mps := 1.0,
       SyncDeviation_M := 0.10, Config := Cfg, Data := Dat);
    ADVANCE_TIME(500000000);
    fb(Reset := FALSE, M1CommandActive := TRUE, M2CommandActive := TRUE, M1Direction := 1, M2Direction := 1,
       M1BrakeCmd := TRUE, M2BrakeCmd := TRUE, M1BrakeApplied := FALSE, M2BrakeApplied := FALSE,
       M1Position_M := 0.5, M2Position_M := 0.5, M1Speed_Mps := 1.0, M2Speed_Mps := 1.0,
       SyncDeviation_M := 0.10, Config := Cfg, Data := Dat);
    ADVANCE_TIME(500000000);
    fb(Reset := FALSE, M1CommandActive := TRUE, M2CommandActive := TRUE, M1Direction := 1, M2Direction := 1,
       M1BrakeCmd := TRUE, M2BrakeCmd := TRUE, M1BrakeApplied := FALSE, M2BrakeApplied := FALSE,
       M1Position_M := 1.0, M2Position_M := 1.0, M1Speed_Mps := 1.0, M2Speed_Mps := 1.0,
       SyncDeviation_M := 0.10, Config := Cfg, Data := Dat);
    ADVANCE_TIME(500000000);
    fb(Reset := FALSE, M1CommandActive := TRUE, M2CommandActive := TRUE, M1Direction := 1, M2Direction := 1,
       M1BrakeCmd := TRUE, M2BrakeCmd := TRUE, M1BrakeApplied := FALSE, M2BrakeApplied := FALSE,
       M1Position_M := 1.5, M2Position_M := 1.5, M1Speed_Mps := 1.0, M2Speed_Mps := 1.0,
       SyncDeviation_M := 0.10, Config := Cfg, Data := Dat);
    ADVANCE_TIME(500000000);
    fb(Reset := FALSE, M1CommandActive := FALSE, M2CommandActive := FALSE, M1Direction := 1, M2Direction := 1,
       M1BrakeCmd := FALSE, M2BrakeCmd := FALSE, M1BrakeApplied := TRUE, M2BrakeApplied := TRUE,
       M1Position_M := 2.0, M2Position_M := 2.0, M1Speed_Mps := 0.0, M2Speed_Mps := 0.0,
       SyncDeviation_M := 0.0, Config := Cfg, Data := Dat);
    ADVANCE_TIME(10000000);
    fb(Reset := FALSE, M1CommandActive := FALSE, M2CommandActive := FALSE, M1Direction := 1, M2Direction := 1,
       M1BrakeCmd := FALSE, M2BrakeCmd := FALSE, M1BrakeApplied := TRUE, M2BrakeApplied := TRUE,
       M1Position_M := 2.0, M2Position_M := 2.0, M1Speed_Mps := 0.0, M2Speed_Mps := 0.0,
       SyncDeviation_M := 0.0, Config := Cfg, Data := Dat);
    ASSERT_TRUE(fb.SymmetryValid, 'Cycle complet qualifie puis arrete -> mesure valide');
    ASSERT_TRUE(fb.SymmetryOk, 'M1 et M2 identiques -> tous les ecarts sous les seuils');
END_TEST

TEST 'TC-P10-T181-18b Reset remet les mesures a zero'
    Cfg.MinimumCommandTime_Ms := 300;
    Cfg.MinimumSpeed_Mps := 0.05;
    Cfg.DeltaStartDelay_Ms := 100; Cfg.DeltaBrakeReleaseTime_Ms := 100;
    Cfg.DeltaBrakeApplyTime_Ms := 100; Cfg.DeltaStopDistance_Mm := 100;
    Cfg.DeltaStopTime_Ms := 200;
    fb(Reset := TRUE, M1CommandActive := FALSE, M2CommandActive := FALSE, M1Direction := 0, M2Direction := 0,
       M1BrakeCmd := FALSE, M2BrakeCmd := FALSE, M1BrakeApplied := TRUE, M2BrakeApplied := TRUE,
       M1Position_M := 0.0, M2Position_M := 0.0, M1Speed_Mps := 0.0, M2Speed_Mps := 0.0,
       SyncDeviation_M := 0.0, Config := Cfg, Data := Dat);
    fb(Reset := FALSE, M1CommandActive := TRUE, M2CommandActive := TRUE, M1Direction := 1, M2Direction := 1,
       M1BrakeCmd := TRUE, M2BrakeCmd := TRUE, M1BrakeApplied := FALSE, M2BrakeApplied := FALSE,
       M1Position_M := 0.0, M2Position_M := 0.0, M1Speed_Mps := 1.0, M2Speed_Mps := 1.0,
       SyncDeviation_M := 0.40, Config := Cfg, Data := Dat);
    ADVANCE_TIME(600000000);
    fb(Reset := FALSE, M1CommandActive := TRUE, M2CommandActive := TRUE, M1Direction := 1, M2Direction := 1,
       M1BrakeCmd := TRUE, M2BrakeCmd := TRUE, M1BrakeApplied := FALSE, M2BrakeApplied := FALSE,
       M1Position_M := 0.6, M2Position_M := 0.6, M1Speed_Mps := 1.0, M2Speed_Mps := 1.0,
       SyncDeviation_M := 0.40, Config := Cfg, Data := Dat);
    ADVANCE_TIME(600000000);
    fb(Reset := FALSE, M1CommandActive := TRUE, M2CommandActive := TRUE, M1Direction := 1, M2Direction := 1,
       M1BrakeCmd := TRUE, M2BrakeCmd := TRUE, M1BrakeApplied := FALSE, M2BrakeApplied := FALSE,
       M1Position_M := 1.2, M2Position_M := 1.2, M1Speed_Mps := 1.0, M2Speed_Mps := 1.0,
       SyncDeviation_M := 0.40, Config := Cfg, Data := Dat);
    fb(Reset := TRUE, M1CommandActive := FALSE, M2CommandActive := FALSE, M1Direction := 0, M2Direction := 0,
       M1BrakeCmd := FALSE, M2BrakeCmd := FALSE, M1BrakeApplied := TRUE, M2BrakeApplied := TRUE,
       M1Position_M := 0.0, M2Position_M := 0.0, M1Speed_Mps := 0.0, M2Speed_Mps := 0.0,
       SyncDeviation_M := 0.0, Config := Cfg, Data := Dat);
    ASSERT_EQ(Dat.DeltaStartDelay_Ms, 0, 'Reset -> DeltaStartDelay_Ms remis a 0');
    ASSERT_FALSE(Dat.MaxSyncDeviation_M > 0.0, 'Reset -> MaxSyncDeviation_M remis a 0');
END_TEST

TEST 'TC-P10-T181-18c Non qualifie si un seul treuil commande'
    Cfg.MinimumCommandTime_Ms := 300;
    Cfg.MinimumSpeed_Mps := 0.05;
    Cfg.DeltaStartDelay_Ms := 100; Cfg.DeltaBrakeReleaseTime_Ms := 100;
    Cfg.DeltaBrakeApplyTime_Ms := 100; Cfg.DeltaStopDistance_Mm := 100;
    Cfg.DeltaStopTime_Ms := 200;
    fb(Reset := TRUE, M1CommandActive := FALSE, M2CommandActive := FALSE, M1Direction := 0, M2Direction := 0,
       M1BrakeCmd := FALSE, M2BrakeCmd := FALSE, M1BrakeApplied := TRUE, M2BrakeApplied := TRUE,
       M1Position_M := 0.0, M2Position_M := 0.0, M1Speed_Mps := 0.0, M2Speed_Mps := 0.0,
       SyncDeviation_M := 0.0, Config := Cfg, Data := Dat);
    fb(Reset := FALSE, M1CommandActive := TRUE, M2CommandActive := FALSE, M1Direction := 1, M2Direction := 0,
       M1BrakeCmd := TRUE, M2BrakeCmd := FALSE, M1BrakeApplied := FALSE, M2BrakeApplied := TRUE,
       M1Position_M := 0.0, M2Position_M := 0.0, M1Speed_Mps := 1.0, M2Speed_Mps := 0.0,
       SyncDeviation_M := 0.30, Config := Cfg, Data := Dat);
    ADVANCE_TIME(1500000000);
    fb(Reset := FALSE, M1CommandActive := TRUE, M2CommandActive := FALSE, M1Direction := 1, M2Direction := 0,
       M1BrakeCmd := TRUE, M2BrakeCmd := FALSE, M1BrakeApplied := FALSE, M2BrakeApplied := TRUE,
       M1Position_M := 1.5, M2Position_M := 0.0, M1Speed_Mps := 1.0, M2Speed_Mps := 0.0,
       SyncDeviation_M := 0.30, Config := Cfg, Data := Dat);
    ASSERT_FALSE(fb.SymmetryValid, 'Un seul treuil commande -> jamais qualifie');
END_TEST

(* ---- FB_WinchLoadEstimator_test.st ---- *)
(* =======================================================================
   test_fb_winchloadestimator.st — T181-18 D11 : macro TC FB_WinchLoadEstimator
   Estimateur informatif (aucune action securite). Couvre : gate, classement
   de vitesse par bande + hysteresis, direction montee/descente, validation table.
   (La lecture de la matrice 5x5 elle-meme n'est pas asserted ici : passthrough,
   et le harnais STruCpp ne supporte pas l'indexation [i][j] d'un ARRAY OF ARRAY.)
   ======================================================================= *)

SETUP
VAR
    fb  : FB_WinchLoadEstimator;
    Spd : ST_fbWinchLoadEstimator_SpeedCfg;
    Tbl : ST_fbWinchLoadEstimator_Table;
END_VAR
END_SETUP

TEST 'TC-P10-T181-18a Gate : Enable FALSE -> sorties neutres'
    Spd.MaxMeasuredSpeedMps := 2.0;
    Spd.SpeedBandMaxMps[1] := 0.4; Spd.SpeedBandMaxMps[2] := 0.8; Spd.SpeedBandMaxMps[3] := 1.2;
    Spd.SpeedBandMaxMps[4] := 1.6; Spd.SpeedBandMaxMps[5] := 2.0;
    Spd.SpeedBandHysteresisMps := 0.05;
    fb(Enable := FALSE, PowerContactorEngaged := TRUE, ActiveSpeedStep := 3,
       MeasuredSpeedMps := 0.5, MeasuredSpeedSignedMps := 0.5,
       SpeedConfig := Spd, LoadTable := Tbl);
    ASSERT_FALSE(fb.Ready, 'Enable FALSE -> Ready FALSE');
    ASSERT_EQ(fb.SpeedBand, 0, 'Enable FALSE -> SpeedBand 0');
    ASSERT_EQ(fb.EstimatedLoadPct, 0.0, 'Enable FALSE -> estimation 0');
END_TEST

TEST 'TC-P10-T181-18b Classement vitesse : 0.5 m/s -> bande 2, montee'
    Spd.MaxMeasuredSpeedMps := 2.0;
    Spd.SpeedBandMaxMps[1] := 0.4; Spd.SpeedBandMaxMps[2] := 0.8; Spd.SpeedBandMaxMps[3] := 1.2;
    Spd.SpeedBandMaxMps[4] := 1.6; Spd.SpeedBandMaxMps[5] := 2.0;
    Spd.SpeedBandHysteresisMps := 0.05;
    Tbl.IsConfigured := TRUE;
    fb(Enable := TRUE, PowerContactorEngaged := TRUE, ActiveSpeedStep := 2,
       MeasuredSpeedMps := 0.5, MeasuredSpeedSignedMps := 0.5,
       SpeedConfig := Spd, LoadTable := Tbl);
    ASSERT_EQ(fb.SpeedBand, 2, 'Vitesse 0.5 m/s (entre 0.4 et 0.8) -> bande 2');
    ASSERT_TRUE(fb.Ascending, 'Vitesse signee positive -> montee');
    ASSERT_TRUE(fb.Configured, 'Table validee -> Configured TRUE');
    ASSERT_TRUE(fb.Ready, 'Nominal -> Ready TRUE');
END_TEST

TEST 'TC-P10-T181-18c Classement vitesse : 1.5 m/s -> bande 4'
    Spd.MaxMeasuredSpeedMps := 2.0;
    Spd.SpeedBandMaxMps[1] := 0.4; Spd.SpeedBandMaxMps[2] := 0.8; Spd.SpeedBandMaxMps[3] := 1.2;
    Spd.SpeedBandMaxMps[4] := 1.6; Spd.SpeedBandMaxMps[5] := 2.0;
    Spd.SpeedBandHysteresisMps := 0.05;
    fb(Enable := TRUE, PowerContactorEngaged := TRUE, ActiveSpeedStep := 4,
       MeasuredSpeedMps := 1.5, MeasuredSpeedSignedMps := 1.5,
       SpeedConfig := Spd, LoadTable := Tbl);
    ASSERT_EQ(fb.SpeedBand, 4, 'Vitesse 1.5 m/s (entre 1.2 et 1.6) -> bande 4');
END_TEST

TEST 'TC-P10-T181-18d Descente : aucune estimation de charge'
    Spd.MaxMeasuredSpeedMps := 2.0;
    Spd.SpeedBandMaxMps[1] := 0.4; Spd.SpeedBandMaxMps[2] := 0.8; Spd.SpeedBandMaxMps[3] := 1.2;
    Spd.SpeedBandMaxMps[4] := 1.6; Spd.SpeedBandMaxMps[5] := 2.0;
    Spd.SpeedBandHysteresisMps := 0.05;
    Tbl.IsConfigured := TRUE;
    fb(Enable := TRUE, PowerContactorEngaged := TRUE, ActiveSpeedStep := 2,
       MeasuredSpeedMps := 0.5, MeasuredSpeedSignedMps := -0.5,
       SpeedConfig := Spd, LoadTable := Tbl);
    ASSERT_FALSE(fb.Ascending, 'Vitesse signee negative -> descente');
    ASSERT_EQ(fb.EstimatedLoadPct, 0.0, 'Descente : estimation non produite');
END_TEST

TEST 'TC-P10-T181-18e Vitesse mesuree negative -> defaut latche, bande 0'
    Spd.MaxMeasuredSpeedMps := 2.0;
    Spd.SpeedBandMaxMps[1] := 0.4; Spd.SpeedBandMaxMps[2] := 0.8; Spd.SpeedBandMaxMps[3] := 1.2;
    Spd.SpeedBandMaxMps[4] := 1.6; Spd.SpeedBandMaxMps[5] := 2.0;
    Spd.SpeedBandHysteresisMps := 0.05;
    fb(Enable := TRUE, PowerContactorEngaged := TRUE, ActiveSpeedStep := 2,
       MeasuredSpeedMps := -0.1, MeasuredSpeedSignedMps := -0.1,
       SpeedConfig := Spd, LoadTable := Tbl);
    ASSERT_EQ(fb.SpeedBand, 0, 'Vitesse mesuree < 0 -> bande 0');
    (* Le socle latche la cause au scan suivant (Active pose apres l'appel FB_FaultCore). *)
    fb(Enable := TRUE, PowerContactorEngaged := TRUE, ActiveSpeedStep := 2,
       MeasuredSpeedMps := -0.1, MeasuredSpeedSignedMps := -0.1,
       SpeedConfig := Spd, LoadTable := Tbl);
    ASSERT_TRUE(fb.Fault.Latched, 'Vitesse mesuree < 0 -> defaut latche');
END_TEST
